(* IEC 61131-3 sources: deprecated-refusr-repo/GP/Main/samples (part 20) *)

(* ---- RND-EXPR_cribs-hyena-lilts.st ---- *)
(*
This code implements a randomly grown symbolic expression:

IN28 & IN39

*)

FUNCTION_BLOCK F_CollectInput
  VAR_IN_OUT
      Data : ARRAY[1..50] OF BOOL;
  END_VAR
  VAR_INPUT
      TICK  : BOOL := 0;
      IN1   : BOOL := 0;
      IN2   : BOOL := 0;
      IN3   : BOOL := 0;
      IN4   : BOOL := 0;
      IN5   : BOOL := 0;
      RESET : BOOL := FALSE;
  END_VAR
  VAR_OUTPUT
      Finished : BOOL;
  END_VAR
  VAR
      j    : USINT := 1;
      tock : BOOL  := 0;
  END_VAR
  IF NOT RESET AND tock = NOT TICK THEN
      Data[j]   := IN1;
      Data[j+1] := IN2;
      Data[j+2] := IN3;
      Data[j+3] := IN4;
      Data[j+4] := IN5;
      j := j + 5;
      tock := TICK;
  ELSE
      j := 1;
      tock := 0;
  END_IF;
  Finished := (j > 50);
END_FUNCTION_BLOCK

PROGRAM Boiler
  VAR
    Data  : ARRAY[1..50] OF BOOL;
    Ready : BOOL;
    CollectInput : F_CollectInput;
  END_VAR
  VAR
    TICK     AT %IX1.0 : BOOL;
    IN1      AT %IX0.3 : BOOL;
    IN2      AT %IX0.4 : BOOL;
    IN3      AT %IX0.5 : BOOL;
    IN4      AT %IX0.6 : BOOL;
    IN5      AT %IX0.7 : BOOL;
    OutReady AT %QX0.0 : BOOL := FALSE;
    FeedNext AT %QX0.1 : BOOL := FALSE;
    Out      AT %QX0.2 : BOOL;
  END_VAR
  CollectInput(TICK:=TICK, IN1:=IN1, IN2:=IN2, IN3:=IN3, IN4:=IN4, IN5:=IN5);
  Ready := CollectInput.Finished;
  FeedNext := 1;
  IF Ready THEN
    Out := (Data[28] AND Data[39]);
    OutReady := 1;
    CollectInput(RESET:=TRUE);
  END_IF;
END_PROGRAM

CONFIGURATION Config0
  RESOURCE Res0 ON PLC
    TASK task0(INTERVAL := T#20ms,PRIORITY := 0);
    PROGRAM instance0 WITH task0 : Boiler;
  END_RESOURCE
END_CONFIGURATION

(* ---- RND-EXPR_culls-boxes-teats.st ---- *)
(*
This code implements a randomly grown symbolic expression:

xor(xor(xor(xor(!((IN48 | (xor(xor(!(!(IN48)), !(!(xor(xor(IN15 & IN37, IN27 & IN43), xor(xor(IN10, IN50), IN49))))), !((IN7 & (xor(xor(IN34, IN29), IN41))) | ((IN34 & IN45) | (!(IN2))))))) & IN16), IN31), IN38), (IN16 | IN47) & IN28), (((!(IN20)) | ((xor(xor(xor(xor(((IN39 | IN35) | (IN9 & IN43)) & IN46, !((!(IN46)) | (xor(xor(IN5, IN34), IN46)))), (!(IN19 | IN49)) | (!(!(IN22)))), xor(xor(IN13, IN22), ((!(IN35)) & (xor(xor(IN2, IN40), IN38))) & IN43)), IN29)) | (xor(xor(!(!(xor(xor(IN8 | IN20, IN6 | IN40), xor(xor(IN12, IN18), IN33)))), !(((!(IN34)) & IN30) | ((!(IN31)) & (IN36 & IN6)))), (!(IN35)) & true)))) & ((((IN17 | (!(!(IN26 | IN42)))) | (xor(xor(IN44, ((xor(xor(IN13, IN3), IN47)) | (xor(xor(IN10, IN45), IN26))) & (xor(xor(!(IN3), IN34 | true), !(IN45)))), !(IN7 | IN35)))) & ((!(!(xor(xor(IN41 & IN25, xor(xor(IN10, IN9), IN48)), IN39)))) | (xor(xor(((xor(xor(IN22, IN35), IN30)) | (IN30 & IN45)) & ((IN24 | IN15) | IN48), !((xor(xor(IN16, IN5), IN23)) | (!(IN4)))), !((xor(xor(IN38, IN16), IN14)) | IN41))))) | ((IN27 & IN46) & ((xor(xor(!(!(xor(xor(IN29, IN24), IN24))), ((IN29 & IN32) & (IN36 | IN47)) | IN15), !(xor(xor(IN45, IN47 | IN29), xor(false, IN9))))) & (xor(xor(xor(xor((xor(xor(IN29, IN4), IN8)) & (!(IN27)), (xor(xor(IN24, IN23), IN10)) | IN19), (IN35 & IN15) | IN20), IN4 & ((!(IN9)) | (xor(xor(IN12, IN15), IN37)))), !(!(IN3)))))))) & (IN27 | IN9))

*)

FUNCTION_BLOCK F_CollectInput
  VAR_IN_OUT
      Data : ARRAY[1..50] OF BOOL;
  END_VAR
  VAR_INPUT
      TICK  : BOOL := 0;
      IN1   : BOOL := 0;
      IN2   : BOOL := 0;
      IN3   : BOOL := 0;
      IN4   : BOOL := 0;
      IN5   : BOOL := 0;
      RESET : BOOL := FALSE;
  END_VAR
  VAR_OUTPUT
      Finished : BOOL;
  END_VAR
  VAR
      j    : USINT := 1;
      tock : BOOL  := 0;
  END_VAR
  IF NOT RESET AND tock = NOT TICK THEN
      Data[j]   := IN1;
      Data[j+1] := IN2;
      Data[j+2] := IN3;
      Data[j+3] := IN4;
      Data[j+4] := IN5;
      j := j + 5;
      tock := TICK;
  ELSE
      j := 1;
      tock := 0;
  END_IF;
  Finished := (j > 50);
END_FUNCTION_BLOCK

PROGRAM Boiler
  VAR
    Data  : ARRAY[1..50] OF BOOL;
    Ready : BOOL;
    CollectInput : F_CollectInput;
  END_VAR
  VAR
    TICK     AT %IX1.0 : BOOL;
    IN1      AT %IX0.3 : BOOL;
    IN2      AT %IX0.4 : BOOL;
    IN3      AT %IX0.5 : BOOL;
    IN4      AT %IX0.6 : BOOL;
    IN5      AT %IX0.7 : BOOL;
    OutReady AT %QX0.0 : BOOL := FALSE;
    FeedNext AT %QX0.1 : BOOL := FALSE;
    Out      AT %QX0.2 : BOOL;
  END_VAR
  CollectInput(TICK:=TICK, IN1:=IN1, IN2:=IN2, IN3:=IN3, IN4:=IN4, IN5:=IN5);
  Ready := CollectInput.Finished;
  FeedNext := 1;
  IF Ready THEN
    Out := (((((NOT ((Data[48] OR (((NOT (NOT Data[48])) XOR (NOT (NOT (((Data[15] AND Data[37]) XOR (Data[27] AND Data[43])) XOR ((Data[10] XOR Data[50]) XOR Data[49]))))) XOR (NOT ((Data[7] AND ((Data[34] XOR Data[29]) XOR Data[41])) OR ((Data[34] AND Data[45]) OR (NOT Data[2])))))) AND Data[16])) XOR Data[31]) XOR Data[38]) XOR ((Data[16] OR Data[47]) AND Data[28])) XOR ((((NOT Data[20]) OR ((((((((Data[39] OR Data[35]) OR (Data[9] AND Data[43])) AND Data[46]) XOR (NOT ((NOT Data[46]) OR ((Data[5] XOR Data[34]) XOR Data[46])))) XOR ((NOT (Data[19] OR Data[49])) OR (NOT (NOT Data[22])))) XOR ((Data[13] XOR Data[22]) XOR (((NOT Data[35]) AND ((Data[2] XOR Data[40]) XOR Data[38])) AND Data[43]))) XOR Data[29]) OR (((NOT (NOT (((Data[8] OR Data[20]) XOR (Data[6] OR Data[40])) XOR ((Data[12] XOR Data[18]) XOR Data[33])))) XOR (NOT (((NOT Data[34]) AND Data[30]) OR ((NOT Data[31]) AND (Data[36] AND Data[6]))))) XOR ((NOT Data[35]) AND TRUE)))) AND ((((Data[17] OR (NOT (NOT (Data[26] OR Data[42])))) OR ((Data[44] XOR ((((Data[13] XOR Data[3]) XOR Data[47]) OR ((Data[10] XOR Data[45]) XOR Data[26])) AND (((NOT Data[3]) XOR (Data[34] OR TRUE)) XOR (NOT Data[45])))) XOR (NOT (Data[7] OR Data[35])))) AND ((NOT (NOT (((Data[41] AND Data[25]) XOR ((Data[10] XOR Data[9]) XOR Data[48])) XOR Data[39]))) OR ((((((Data[22] XOR Data[35]) XOR Data[30]) OR (Data[30] AND Data[45])) AND ((Data[24] OR Data[15]) OR Data[48])) XOR (NOT (((Data[16] XOR Data[5]) XOR Data[23]) OR (NOT Data[4])))) XOR (NOT (((Data[38] XOR Data[16]) XOR Data[14]) OR Data[41]))))) OR ((Data[27] AND Data[46]) AND ((((NOT (NOT ((Data[29] XOR Data[24]) XOR Data[24]))) XOR (((Data[29] AND Data[32]) AND (Data[36] OR Data[47])) OR Data[15])) XOR (NOT ((Data[45] XOR (Data[47] OR Data[29])) XOR (FALSE XOR Data[9])))) AND (((((((Data[29] XOR Data[4]) XOR Data[8]) AND (NOT Data[27])) XOR (((Data[24] XOR Data[23]) XOR Data[10]) OR Data[19])) XOR ((Data[35] AND Data[15]) OR Data[20])) XOR (Data[4] AND ((NOT Data[9]) OR ((Data[12] XOR Data[15]) XOR Data[37])))) XOR (NOT (NOT Data[3]))))))) AND (Data[27] OR Data[9])));
    OutReady := 1;
    CollectInput(RESET:=TRUE);
  END_IF;
END_PROGRAM

CONFIGURATION Config0
  RESOURCE Res0 ON PLC
    TASK task0(INTERVAL := T#20ms,PRIORITY := 0);
    PROGRAM instance0 WITH task0 : Boiler;
  END_RESOURCE
END_CONFIGURATION

(* ---- RND-EXPR_datum-botch-beams.st ---- *)
(*
This code implements a randomly grown symbolic expression:

(((xor(xor((xor(xor(xor(xor(IN19, (!(IN48 | IN21)) & (!(xor(xor(IN30, IN18), IN5)))), IN21), ((xor(xor(IN23 | IN7, IN44 | IN43), IN28 & IN45)) & ((!(IN4)) | (IN37 | IN4))) | (xor(xor((IN10 | IN19) | (IN27 & IN18), IN45), !(IN41)))), IN21)) & ((((IN36 | false) | ((!(IN22)) | (xor(xor(IN17, IN20), IN45)))) | (((xor(xor(IN40, IN49), IN35)) & (!(IN19))) & (xor(xor(xor(xor(IN32, IN22), IN46), !(IN2)), xor(xor(IN46, IN23), IN28))))) | ((((IN7 & IN47) & (IN5 & IN32)) & ((IN29 | IN13) | (true & IN42))) & ((true & (IN8 & IN29)) & (xor(xor(!(IN46), !(IN24)), xor(xor(IN6, IN16), IN4)))))), (((!(!(IN20 | IN46))) | (!(xor(xor(!(IN16), xor(xor(IN12, IN9), IN4)), IN31 | IN40)))) & IN49) & (xor(xor(IN41, (xor(xor((xor(xor(true, IN18), false)) & (xor(xor(IN10, IN15), IN4)), (!(IN14)) & IN12), (IN43 | IN32) & IN32)) & (IN31 | ((xor(xor(IN22, true), IN17)) | (xor(xor(IN49, IN20), false))))), xor(xor(!(IN45), IN46), IN2 | (xor(xor(IN11, IN2 & IN18), IN43 | IN11)))))), IN11)) | IN13) | (xor(xor(xor(xor((!((!((IN29 | IN7) & (IN48 | IN42))) | IN20)) | (!(IN21)), (xor(xor(xor(xor(xor(xor((xor(xor(IN1, IN10), IN29)) | (IN2 & IN25), xor(xor(xor(xor(IN34, IN6), IN25), IN41 & IN10), IN36 & IN25)), (IN6 & IN20) | (IN47 | IN26)), IN7), !((IN43 & IN25) | (xor(xor(IN44, IN44), IN30)))), IN15 | (IN8 & (xor(xor(xor(xor(IN3, IN16), IN33), IN3 & IN40), !(IN40))))), IN31 & IN19)) & (IN27 & (!(IN47 & (xor(xor(IN5, IN38 & IN40), IN30)))))), xor(xor(((!(!(IN24))) & (xor(xor(IN30, IN2), xor(xor(xor(xor(IN38, true), IN8), IN33 & IN9), xor(xor(IN49, IN40), IN43))))) & (((true & (xor(xor(IN49, IN36), IN7))) | ((!(IN21)) | (IN4 & IN40))) & IN47), ((((IN13 | IN3) & IN30) & (xor(xor(IN3 & IN14, !(IN41)), !(IN22)))) & ((!(IN33 | IN21)) | (!(IN18 & IN42)))) | (xor(xor((xor(xor(!(IN37), IN49 | IN14), IN42)) & (!(IN1 & IN30)), ((!(IN18)) & (xor(xor(IN28, IN28), IN42))) & (IN40 | IN32)), !(IN34 & (xor(xor(IN45, IN21), IN18)))))), xor(xor(!(!(xor(xor(IN48 | IN1, !(IN12)), !(IN27)))), ((xor(xor(IN43 | IN15, IN9 | IN20), xor(xor(IN4, IN4), IN11))) & IN35) & (IN21 | (!(IN13 & IN21)))), ((xor(xor(xor(xor(IN29, IN17), IN6), IN23 | IN2), IN46 | IN28)) & (!(IN42))) | IN9))), xor(xor(IN21, !(!(!(!((xor(xor(IN47, IN29), IN31)) & (IN3 & IN43)))))), (!((xor(xor(!(IN27 | IN39), xor(xor(xor(xor(IN1, IN14), IN16), false | IN8), IN47 | IN1)), xor(xor(IN36 & IN31, !(IN39)), IN44 | IN33))) & ((IN8 | (IN5 | IN34)) & (!(xor(xor(IN12, IN31), IN12)))))) | ((((!(xor(xor(IN45, IN8), IN46))) & IN45) & IN8) | (!(!((IN28 & IN42) & (IN50 | IN35))))))), xor(xor(IN29, !((IN34 | (IN1 | (IN12 & (IN6 | IN15)))) & ((!(!(IN32 & IN18))) & (!(!(IN6 & IN28)))))), ((!(!(IN25))) | (xor(xor(xor(xor(!(IN3 & IN34), xor(xor(IN16 & IN26, !(IN26)), IN17)), (IN33 & IN37) & (!(IN32))), ((IN38 | IN8) & (!(IN19))) | (xor(xor(!(IN29), IN4 | IN21), IN39 & IN36))), (xor(xor(IN41 | IN43, xor(xor(IN32, IN10), IN28)), IN18 & IN1)) | (IN25 & IN34)))) & IN8)))) | IN13

*)

FUNCTION_BLOCK F_CollectInput
  VAR_IN_OUT
      Data : ARRAY[1..50] OF BOOL;
  END_VAR
  VAR_INPUT
      TICK  : BOOL := 0;
      IN1   : BOOL := 0;
      IN2   : BOOL := 0;
      IN3   : BOOL := 0;
      IN4   : BOOL := 0;
      IN5   : BOOL := 0;
      RESET : BOOL := FALSE;
  END_VAR
  VAR_OUTPUT
      Finished : BOOL;
  END_VAR
  VAR
      j    : USINT := 1;
      tock : BOOL  := 0;
  END_VAR
  IF NOT RESET AND tock = NOT TICK THEN
      Data[j]   := IN1;
      Data[j+1] := IN2;
      Data[j+2] := IN3;
      Data[j+3] := IN4;
      Data[j+4] := IN5;
      j := j + 5;
      tock := TICK;
  ELSE
      j := 1;
      tock := 0;
  END_IF;
  Finished := (j > 50);
END_FUNCTION_BLOCK

PROGRAM Boiler
  VAR
    Data  : ARRAY[1..50] OF BOOL;
    Ready : BOOL;
    CollectInput : F_CollectInput;
  END_VAR
  VAR
    TICK     AT %IX1.0 : BOOL;
    IN1      AT %IX0.3 : BOOL;
    IN2      AT %IX0.4 : BOOL;
    IN3      AT %IX0.5 : BOOL;
    IN4      AT %IX0.6 : BOOL;
    IN5      AT %IX0.7 : BOOL;
    OutReady AT %QX0.0 : BOOL := FALSE;
    FeedNext AT %QX0.1 : BOOL := FALSE;
    Out      AT %QX0.2 : BOOL;
  END_VAR
  CollectInput(TICK:=TICK, IN1:=IN1, IN2:=IN2, IN3:=IN3, IN4:=IN4, IN5:=IN5);
  Ready := CollectInput.Finished;
  FeedNext := 1;
  IF Ready THEN
    Out := ((((((((((Data[19] XOR ((NOT (Data[48] OR Data[21])) AND (NOT ((Data[30] XOR Data[18]) XOR Data[5])))) XOR Data[21]) XOR (((((Data[23] OR Data[7]) XOR (Data[44] OR Data[43])) XOR (Data[28] AND Data[45])) AND ((NOT Data[4]) OR (Data[37] OR Data[4]))) OR ((((Data[10] OR Data[19]) OR (Data[27] AND Data[18])) XOR Data[45]) XOR (NOT Data[41])))) XOR Data[21]) AND ((((Data[36] OR FALSE) OR ((NOT Data[22]) OR ((Data[17] XOR Data[20]) XOR Data[45]))) OR ((((Data[40] XOR Data[49]) XOR Data[35]) AND (NOT Data[19])) AND ((((Data[32] XOR Data[22]) XOR Data[46]) XOR (NOT Data[2])) XOR ((Data[46] XOR Data[23]) XOR Data[28])))) OR ((((Data[7] AND Data[47]) AND (Data[5] AND Data[32])) AND ((Data[29] OR Data[13]) OR (TRUE AND Data[42]))) AND ((TRUE AND (Data[8] AND Data[29])) AND (((NOT Data[46]) XOR (NOT Data[24])) XOR ((Data[6] XOR Data[16]) XOR Data[4])))))) XOR ((((NOT (NOT (Data[20] OR Data[46]))) OR (NOT (((NOT Data[16]) XOR ((Data[12] XOR Data[9]) XOR Data[4])) XOR (Data[31] OR Data[40])))) AND Data[49]) AND ((Data[41] XOR ((((((TRUE XOR Data[18]) XOR FALSE) AND ((Data[10] XOR Data[15]) XOR Data[4])) XOR ((NOT Data[14]) AND Data[12])) XOR ((Data[43] OR Data[32]) AND Data[32])) AND (Data[31] OR (((Data[22] XOR TRUE) XOR Data[17]) OR ((Data[49] XOR Data[20]) XOR FALSE))))) XOR (((NOT Data[45]) XOR Data[46]) XOR (Data[2] OR ((Data[11] XOR (Data[2] AND Data[18])) XOR (Data[43] OR Data[11]))))))) XOR Data[11]) OR Data[13]) OR ((((((NOT ((NOT ((Data[29] OR Data[7]) AND (Data[48] OR Data[42]))) OR Data[20])) OR (NOT Data[21])) XOR ((((((((((Data[1] XOR Data[10]) XOR Data[29]) OR (Data[2] AND Data[25])) XOR ((((Data[34] XOR Data[6]) XOR Data[25]) XOR (Data[41] AND Data[10])) XOR (Data[36] AND Data[25]))) XOR ((Data[6] AND Data[20]) OR (Data[47] OR Data[26]))) XOR Data[7]) XOR (NOT ((Data[43] AND Data[25]) OR ((Data[44] XOR Data[44]) XOR Data[30])))) XOR (Data[15] OR (Data[8] AND ((((Data[3] XOR Data[16]) XOR Data[33]) XOR (Data[3] AND Data[40])) XOR (NOT Data[40]))))) XOR (Data[31] AND Data[19])) AND (Data[27] AND (NOT (Data[47] AND ((Data[5] XOR (Data[38] AND Data[40])) XOR Data[30])))))) XOR (((((NOT (NOT Data[24])) AND ((Data[30] XOR Data[2]) XOR ((((Data[38] XOR TRUE) XOR Data[8]) XOR (Data[33] AND Data[9])) XOR ((Data[49] XOR Data[40]) XOR Data[43])))) AND (((TRUE AND ((Data[49] XOR Data[36]) XOR Data[7])) OR ((NOT Data[21]) OR (Data[4] AND Data[40]))) AND Data[47])) XOR (((((Data[13] OR Data[3]) AND Data[30]) AND (((Data[3] AND Data[14]) XOR (NOT Data[41])) XOR (NOT Data[22]))) AND ((NOT (Data[33] OR Data[21])) OR (NOT (Data[18] AND Data[42])))) OR ((((((NOT Data[37]) XOR (Data[49] OR Data[14])) XOR Data[42]) AND (NOT (Data[1] AND Data[30]))) XOR (((NOT Data[18]) AND ((Data[28] XOR Data[28]) XOR Data[42])) AND (Data[40] OR Data[32]))) XOR (NOT (Data[34] AND ((Data[45] XOR Data[21]) XOR Data[18])))))) XOR (((NOT (NOT (((Data[48] OR Data[1]) XOR (NOT Data[12])) XOR (NOT Data[27])))) XOR (((((Data[43] OR Data[15]) XOR (Data[9] OR Data[20])) XOR ((Data[4] XOR Data[4]) XOR Data[11])) AND Data[35]) AND (Data[21] OR (NOT (Data[13] AND Data[21]))))) XOR ((((((Data[29] XOR Data[17]) XOR Data[6]) XOR (Data[23] OR Data[2])) XOR (Data[46] OR Data[28])) AND (NOT Data[42])) OR Data[9])))) XOR ((Data[21] XOR (NOT (NOT (NOT (NOT (((Data[47] XOR Data[29]) XOR Data[31]) AND (Data[3] AND Data[43]))))))) XOR ((NOT ((((NOT (Data[27] OR Data[39])) XOR ((((Data[1] XOR Data[14]) XOR Data[16]) XOR (FALSE OR Data[8])) XOR (Data[47] OR Data[1]))) XOR (((Data[36] AND Data[31]) XOR (NOT Data[39])) XOR (Data[44] OR Data[33]))) AND ((Data[8] OR (Data[5] OR Data[34])) AND (NOT ((Data[12] XOR Data[31]) XOR Data[12]))))) OR ((((NOT ((Data[45] XOR Data[8]) XOR Data[46])) AND Data[45]) AND Data[8]) OR (NOT (NOT ((Data[28] AND Data[42]) AND (Data[50] OR Data[35])))))))) XOR ((Data[29] XOR (NOT ((Data[34] OR (Data[1] OR (Data[12] AND (Data[6] OR Data[15])))) AND ((NOT (NOT (Data[32] AND Data[18]))) AND (NOT (NOT (Data[6] AND Data[28]))))))) XOR (((NOT (NOT Data[25])) OR (((((NOT (Data[3] AND Data[34])) XOR (((Data[16] AND Data[26]) XOR (NOT Data[26])) XOR Data[17])) XOR ((Data[33] AND Data[37]) AND (NOT Data[32]))) XOR (((Data[38] OR Data[8]) AND (NOT Data[19])) OR (((NOT Data[29]) XOR (Data[4] OR Data[21])) XOR (Data[39] AND Data[36])))) XOR ((((Data[41] OR Data[43]) XOR ((Data[32] XOR Data[10]) XOR Data[28])) XOR (Data[18] AND Data[1])) OR (Data[25] AND Data[34])))) AND Data[8])))) OR Data[13]);
    OutReady := 1;
    CollectInput(RESET:=TRUE);
  END_IF;
END_PROGRAM

CONFIGURATION Config0
  RESOURCE Res0 ON PLC
    TASK task0(INTERVAL := T#20ms,PRIORITY := 0);
    PROGRAM instance0 WITH task0 : Boiler;
  END_RESOURCE
END_CONFIGURATION

(* ---- RND-EXPR_didot-crows-snoot.st ---- *)
(*
This code implements a randomly grown symbolic expression:

((((xor(xor(IN5, xor(xor(xor(xor(((IN48 & IN29) | (IN9 | IN16)) & ((!(IN32)) & (xor(xor(IN31, IN7), IN31))), IN21 & (!(!(IN38)))), IN40 & ((IN8 & IN7) & (!(IN26)))), !(xor(xor(!(!(IN18)), xor(xor(IN2 & IN4, xor(xor(IN20, IN39), IN3)), IN20)), !(xor(xor(IN38, IN20), IN30))))), xor(xor(!(IN10), xor(xor(IN9, (!(IN6)) & (true & IN13)), xor(xor(xor(xor(IN27, IN43), false), xor(xor(IN49, IN1), IN26)), !(IN6)))), (!(!(IN27))) | (IN47 & (IN34 & IN35))))), (xor(xor(IN44, (!(!(IN15))) & (xor(xor(IN27 & IN46, IN40 & IN32), !(IN14)))), xor(xor(!(IN46 & IN21), !(!(IN46))), (xor(xor(IN25, IN12), IN13)) | (!(IN50))))) | (IN20 | ((!(xor(xor(IN22, IN46), IN28))) | (!(IN24)))))) & (((((IN24 & (!(IN48))) & (!(IN22))) | (!(!(!(IN24))))) | ((xor(xor((!(IN2)) | (!(IN5)), IN46), xor(xor(IN45 & IN25, IN43), IN43))) & (xor(xor(xor(xor(IN7, !(IN33)), xor(xor(IN3, IN5), IN17)), xor(xor(IN39 & IN18, !(IN8)), IN15 & IN24)), (!(IN38)) | (IN9 | IN17))))) & (xor(xor(IN20 & (xor(xor((IN35 | IN47) & (xor(xor(IN46, IN9), IN16)), IN17), xor(xor(!(IN14), IN31), !(IN44)))), xor(xor((xor(xor(xor(xor(IN38, IN15), IN25), IN36 & IN30), IN7 & IN34)) | (!(xor(xor(IN31, IN21), IN10))), !(xor(xor(xor(xor(IN47, IN11), IN2), IN25 | IN46), IN10))), IN21)), IN45)))) | (xor(xor(IN46 & (IN16 | (!((IN31 & (!(IN12))) & (!(IN31 & IN34))))), IN43 | ((!((!(IN7 | IN36)) | IN29)) & (!((xor(xor(!(IN39), IN7), xor(xor(IN2, IN38), IN16))) | (xor(xor(IN21 & IN38, IN39 | IN14), IN28 & IN3)))))), !(!(!(IN5 | (!(IN5 & IN46)))))))) & IN50) & IN18

*)

FUNCTION_BLOCK F_CollectInput
  VAR_IN_OUT
      Data : ARRAY[1..50] OF BOOL;
  END_VAR
  VAR_INPUT
      TICK  : BOOL := 0;
      IN1   : BOOL := 0;
      IN2   : BOOL := 0;
      IN3   : BOOL := 0;
      IN4   : BOOL := 0;
      IN5   : BOOL := 0;
      RESET : BOOL := FALSE;
  END_VAR
  VAR_OUTPUT
      Finished : BOOL;
  END_VAR
  VAR
      j    : USINT := 1;
      tock : BOOL  := 0;
  END_VAR
  IF NOT RESET AND tock = NOT TICK THEN
      Data[j]   := IN1;
      Data[j+1] := IN2;
      Data[j+2] := IN3;
      Data[j+3] := IN4;
      Data[j+4] := IN5;
      j := j + 5;
      tock := TICK;
  ELSE
      j := 1;
      tock := 0;
  END_IF;
  Finished := (j > 50);
END_FUNCTION_BLOCK

PROGRAM Boiler
  VAR
    Data  : ARRAY[1..50] OF BOOL;
    Ready : BOOL;
    CollectInput : F_CollectInput;
  END_VAR
  VAR
    TICK     AT %IX1.0 : BOOL;
    IN1      AT %IX0.3 : BOOL;
    IN2      AT %IX0.4 : BOOL;
    IN3      AT %IX0.5 : BOOL;
    IN4      AT %IX0.6 : BOOL;
    IN5      AT %IX0.7 : BOOL;
    OutReady AT %QX0.0 : BOOL := FALSE;
    FeedNext AT %QX0.1 : BOOL := FALSE;
    Out      AT %QX0.2 : BOOL;
  END_VAR
  CollectInput(TICK:=TICK, IN1:=IN1, IN2:=IN2, IN3:=IN3, IN4:=IN4, IN5:=IN5);
  Ready := CollectInput.Finished;
  FeedNext := 1;
  IF Ready THEN
    Out := ((((((Data[5] XOR (((((((Data[48] AND Data[29]) OR (Data[9] OR Data[16])) AND ((NOT Data[32]) AND ((Data[31] XOR Data[7]) XOR Data[31]))) XOR (Data[21] AND (NOT (NOT Data[38])))) XOR (Data[40] AND ((Data[8] AND Data[7]) AND (NOT Data[26])))) XOR (NOT (((NOT (NOT Data[18])) XOR (((Data[2] AND Data[4]) XOR ((Data[20] XOR Data[39]) XOR Data[3])) XOR Data[20])) XOR (NOT ((Data[38] XOR Data[20]) XOR Data[30]))))) XOR (((NOT Data[10]) XOR ((Data[9] XOR ((NOT Data[6]) AND (TRUE AND Data[13]))) XOR ((((Data[27] XOR Data[43]) XOR FALSE) XOR ((Data[49] XOR Data[1]) XOR Data[26])) XOR (NOT Data[6])))) XOR ((NOT (NOT Data[27])) OR (Data[47] AND (Data[34] AND Data[35])))))) XOR (((Data[44] XOR ((NOT (NOT Data[15])) AND (((Data[27] AND Data[46]) XOR (Data[40] AND Data[32])) XOR (NOT Data[14])))) XOR (((NOT (Data[46] AND Data[21])) XOR (NOT (NOT Data[46]))) XOR (((Data[25] XOR Data[12]) XOR Data[13]) OR (NOT Data[50])))) OR (Data[20] OR ((NOT ((Data[22] XOR Data[46]) XOR Data[28])) OR (NOT Data[24]))))) AND (((((Data[24] AND (NOT Data[48])) AND (NOT Data[22])) OR (NOT (NOT (NOT Data[24])))) OR (((((NOT Data[2]) OR (NOT Data[5])) XOR Data[46]) XOR (((Data[45] AND Data[25]) XOR Data[43]) XOR Data[43])) AND ((((Data[7] XOR (NOT Data[33])) XOR ((Data[3] XOR Data[5]) XOR Data[17])) XOR (((Data[39] AND Data[18]) XOR (NOT Data[8])) XOR (Data[15] AND Data[24]))) XOR ((NOT Data[38]) OR (Data[9] OR Data[17]))))) AND (((Data[20] AND ((((Data[35] OR Data[47]) AND ((Data[46] XOR Data[9]) XOR Data[16])) XOR Data[17]) XOR (((NOT Data[14]) XOR Data[31]) XOR (NOT Data[44])))) XOR (((((((Data[38] XOR Data[15]) XOR Data[25]) XOR (Data[36] AND Data[30])) XOR (Data[7] AND Data[34])) OR (NOT ((Data[31] XOR Data[21]) XOR Data[10]))) XOR (NOT ((((Data[47] XOR Data[11]) XOR Data[2]) XOR (Data[25] OR Data[46])) XOR Data[10]))) XOR Data[21])) XOR Data[45]))) OR (((Data[46] AND (Data[16] OR (NOT ((Data[31] AND (NOT Data[12])) AND (NOT (Data[31] AND Data[34])))))) XOR (Data[43] OR ((NOT ((NOT (Data[7] OR Data[36])) OR Data[29])) AND (NOT ((((NOT Data[39]) XOR Data[7]) XOR ((Data[2] XOR Data[38]) XOR Data[16])) OR (((Data[21] AND Data[38]) XOR (Data[39] OR Data[14])) XOR (Data[28] AND Data[3]))))))) XOR (NOT (NOT (NOT (Data[5] OR (NOT (Data[5] AND Data[46])))))))) AND Data[50]) AND Data[18]);
    OutReady := 1;
    CollectInput(RESET:=TRUE);
  END_IF;
END_PROGRAM

CONFIGURATION Config0
  RESOURCE Res0 ON PLC
    TASK task0(INTERVAL := T#20ms,PRIORITY := 0);
    PROGRAM instance0 WITH task0 : Boiler;
  END_RESOURCE
END_CONFIGURATION

(* ---- RND-EXPR_dotty-douse-lurer.st ---- *)
(*
This code implements a randomly grown symbolic expression:

xor(xor(!(xor(xor(((xor(xor(IN28, false), (xor(xor((IN5 | IN20) & IN27, (IN25 & IN12) & (!(IN47))), xor(xor(IN14 | IN16, xor(xor(IN17, IN42), IN9)), IN6 | IN50))) | (!(xor(xor(IN20 & IN18, IN41 & false), !(IN41)))))) & (!(!(xor(xor((IN4 | IN22) | (IN4 & IN4), (!(IN31)) & (!(IN11))), !(!(IN25))))))) | (IN22 | (!((((IN15 | IN11) & (IN10 | IN33)) | ((xor(xor(IN28, IN28), IN26)) & (IN10 & IN11))) | IN27))), !(!((xor(xor((xor(xor(IN4 & IN11, xor(xor(IN28, IN40), IN2)), IN2 | IN17)) & (!(IN16)), xor(xor(IN21 | (IN43 | IN19), xor(xor(IN42, IN25 | IN18), IN25 & IN49)), xor(xor(true, IN35 | true), !(IN36)))), (!(IN6 & IN31)) | (!(IN42 & IN48)))) & (xor(xor(IN22, (!(IN30)) | (xor(xor(!(IN11), !(IN42)), IN1 | IN27))), IN7 | ((IN2 | IN23) | (IN30 | IN49))))))), !(IN20 | (IN16 & ((!((IN39 & IN22) & (!(IN7)))) | (!(xor(xor(IN8 | IN15, IN21 | IN44), !(IN2))))))))), IN28), !(!(IN41 | (!(xor(xor(!(xor(xor(xor(xor(IN34 | IN30, IN36), xor(xor(IN31, IN38), IN14)), xor(xor(IN7 & IN44, IN11 & IN13), IN5 & IN15)), !(IN11 & IN10))), (IN14 | false) | IN29), (!(IN47)) & (!((xor(xor(IN17, IN6), IN4)) | (IN47 | IN10)))))))))

*)

FUNCTION_BLOCK F_CollectInput
  VAR_IN_OUT
      Data : ARRAY[1..50] OF BOOL;
  END_VAR
  VAR_INPUT
      TICK  : BOOL := 0;
      IN1   : BOOL := 0;
      IN2   : BOOL := 0;
      IN3   : BOOL := 0;
      IN4   : BOOL := 0;
      IN5   : BOOL := 0;
      RESET : BOOL := FALSE;
  END_VAR
  VAR_OUTPUT
      Finished : BOOL;
  END_VAR
  VAR
      j    : USINT := 1;
      tock : BOOL  := 0;
  END_VAR
  IF NOT RESET AND tock = NOT TICK THEN
      Data[j]   := IN1;
      Data[j+1] := IN2;
      Data[j+2] := IN3;
      Data[j+3] := IN4;
      Data[j+4] := IN5;
      j := j + 5;
      tock := TICK;
  ELSE
      j := 1;
      tock := 0;
  END_IF;
  Finished := (j > 50);
END_FUNCTION_BLOCK

PROGRAM Boiler
  VAR
    Data  : ARRAY[1..50] OF BOOL;
    Ready : BOOL;
    CollectInput : F_CollectInput;
  END_VAR
  VAR
    TICK     AT %IX1.0 : BOOL;
    IN1      AT %IX0.3 : BOOL;
    IN2      AT %IX0.4 : BOOL;
    IN3      AT %IX0.5 : BOOL;
    IN4      AT %IX0.6 : BOOL;
    IN5      AT %IX0.7 : BOOL;
    OutReady AT %QX0.0 : BOOL := FALSE;
    FeedNext AT %QX0.1 : BOOL := FALSE;
    Out      AT %QX0.2 : BOOL;
  END_VAR
  CollectInput(TICK:=TICK, IN1:=IN1, IN2:=IN2, IN3:=IN3, IN4:=IN4, IN5:=IN5);
  Ready := CollectInput.Finished;
  FeedNext := 1;
  IF Ready THEN
    Out := (((NOT ((((((Data[28] XOR FALSE) XOR (((((Data[5] OR Data[20]) AND Data[27]) XOR ((Data[25] AND Data[12]) AND (NOT Data[47]))) XOR (((Data[14] OR Data[16]) XOR ((Data[17] XOR Data[42]) XOR Data[9])) XOR (Data[6] OR Data[50]))) OR (NOT (((Data[20] AND Data[18]) XOR (Data[41] AND FALSE)) XOR (NOT Data[41]))))) AND (NOT (NOT ((((Data[4] OR Data[22]) OR (Data[4] AND Data[4])) XOR ((NOT Data[31]) AND (NOT Data[11]))) XOR (NOT (NOT Data[25])))))) OR (Data[22] OR (NOT ((((Data[15] OR Data[11]) AND (Data[10] OR Data[33])) OR (((Data[28] XOR Data[28]) XOR Data[26]) AND (Data[10] AND Data[11]))) OR Data[27])))) XOR (NOT (NOT (((((((Data[4] AND Data[11]) XOR ((Data[28] XOR Data[40]) XOR Data[2])) XOR (Data[2] OR Data[17])) AND (NOT Data[16])) XOR (((Data[21] OR (Data[43] OR Data[19])) XOR ((Data[42] XOR (Data[25] OR Data[18])) XOR (Data[25] AND Data[49]))) XOR ((TRUE XOR (Data[35] OR TRUE)) XOR (NOT Data[36])))) XOR ((NOT (Data[6] AND Data[31])) OR (NOT (Data[42] AND Data[48])))) AND ((Data[22] XOR ((NOT Data[30]) OR (((NOT Data[11]) XOR (NOT Data[42])) XOR (Data[1] OR Data[27])))) XOR (Data[7] OR ((Data[2] OR Data[23]) OR (Data[30] OR Data[49])))))))) XOR (NOT (Data[20] OR (Data[16] AND ((NOT ((Data[39] AND Data[22]) AND (NOT Data[7]))) OR (NOT (((Data[8] OR Data[15]) XOR (Data[21] OR Data[44])) XOR (NOT Data[2]))))))))) XOR Data[28]) XOR (NOT (NOT (Data[41] OR (NOT (((NOT (((((Data[34] OR Data[30]) XOR Data[36]) XOR ((Data[31] XOR Data[38]) XOR Data[14])) XOR (((Data[7] AND Data[44]) XOR (Data[11] AND Data[13])) XOR (Data[5] AND Data[15]))) XOR (NOT (Data[11] AND Data[10])))) XOR ((Data[14] OR FALSE) OR Data[29])) XOR ((NOT Data[47]) AND (NOT (((Data[17] XOR Data[6]) XOR Data[4]) OR (Data[47] OR Data[10]))))))))));
    OutReady := 1;
    CollectInput(RESET:=TRUE);
  END_IF;
END_PROGRAM

CONFIGURATION Config0
  RESOURCE Res0 ON PLC
    TASK task0(INTERVAL := T#20ms,PRIORITY := 0);
    PROGRAM instance0 WITH task0 : Boiler;
  END_RESOURCE
END_CONFIGURATION

(* ---- RND-EXPR_doxie-capos-donna.st ---- *)
(*
This code implements a randomly grown symbolic expression:

!(!(xor(xor(IN7 | ((((!(xor(xor(IN46, IN6 & IN48), IN36 | IN35))) | (!((xor(xor(IN26, IN22), IN45)) | (IN5 | true)))) | (!(((IN23 & IN25) & IN7) | (xor(xor(xor(xor(IN6, IN4), true), xor(xor(IN2, IN20), IN9)), xor(xor(IN4, IN11), IN36)))))) & (!(IN23))), IN8), ((!((((IN36 & IN24) | (IN45 | IN45)) | ((!(IN8)) | (!(IN23)))) & ((xor(xor(xor(xor(IN41, IN42), IN5), xor(xor(IN5, IN3), IN41)), xor(xor(IN20, IN39), true))) & (xor(xor(!(IN12), IN47 & false), IN14 & IN23))))) | (xor(xor((!(IN3)) & (((xor(xor(IN24, IN43), IN28)) | (!(IN10))) & (!(IN22 | IN28))), IN16), (xor(xor(IN1, IN1), (IN16 & true) | (IN40 | IN50))) & (!(IN39 & (IN8 & IN8)))))) | IN3)))

*)

FUNCTION_BLOCK F_CollectInput
  VAR_IN_OUT
      Data : ARRAY[1..50] OF BOOL;
  END_VAR
  VAR_INPUT
      TICK  : BOOL := 0;
      IN1   : BOOL := 0;
      IN2   : BOOL := 0;
      IN3   : BOOL := 0;
      IN4   : BOOL := 0;
      IN5   : BOOL := 0;
      RESET : BOOL := FALSE;
  END_VAR
  VAR_OUTPUT
      Finished : BOOL;
  END_VAR
  VAR
      j    : USINT := 1;
      tock : BOOL  := 0;
  END_VAR
  IF NOT RESET AND tock = NOT TICK THEN
      Data[j]   := IN1;
      Data[j+1] := IN2;
      Data[j+2] := IN3;
      Data[j+3] := IN4;
      Data[j+4] := IN5;
      j := j + 5;
      tock := TICK;
  ELSE
      j := 1;
      tock := 0;
  END_IF;
  Finished := (j > 50);
END_FUNCTION_BLOCK

PROGRAM Boiler
  VAR
    Data  : ARRAY[1..50] OF BOOL;
    Ready : BOOL;
    CollectInput : F_CollectInput;
  END_VAR
  VAR
    TICK     AT %IX1.0 : BOOL;
    IN1      AT %IX0.3 : BOOL;
    IN2      AT %IX0.4 : BOOL;
    IN3      AT %IX0.5 : BOOL;
    IN4      AT %IX0.6 : BOOL;
    IN5      AT %IX0.7 : BOOL;
    OutReady AT %QX0.0 : BOOL := FALSE;
    FeedNext AT %QX0.1 : BOOL := FALSE;
    Out      AT %QX0.2 : BOOL;
  END_VAR
  CollectInput(TICK:=TICK, IN1:=IN1, IN2:=IN2, IN3:=IN3, IN4:=IN4, IN5:=IN5);
  Ready := CollectInput.Finished;
  FeedNext := 1;
  IF Ready THEN
    Out := (NOT (NOT (((Data[7] OR ((((NOT ((Data[46] XOR (Data[6] AND Data[48])) XOR (Data[36] OR Data[35]))) OR (NOT (((Data[26] XOR Data[22]) XOR Data[45]) OR (Data[5] OR TRUE)))) OR (NOT (((Data[23] AND Data[25]) AND Data[7]) OR ((((Data[6] XOR Data[4]) XOR TRUE) XOR ((Data[2] XOR Data[20]) XOR Data[9])) XOR ((Data[4] XOR Data[11]) XOR Data[36]))))) AND (NOT Data[23]))) XOR Data[8]) XOR (((NOT ((((Data[36] AND Data[24]) OR (Data[45] OR Data[45])) OR ((NOT Data[8]) OR (NOT Data[23]))) AND (((((Data[41] XOR Data[42]) XOR Data[5]) XOR ((Data[5] XOR Data[3]) XOR Data[41])) XOR ((Data[20] XOR Data[39]) XOR TRUE)) AND (((NOT Data[12]) XOR (Data[47] AND FALSE)) XOR (Data[14] AND Data[23]))))) OR ((((NOT Data[3]) AND ((((Data[24] XOR Data[43]) XOR Data[28]) OR (NOT Data[10])) AND (NOT (Data[22] OR Data[28])))) XOR Data[16]) XOR (((Data[1] XOR Data[1]) XOR ((Data[16] AND TRUE) OR (Data[40] OR Data[50]))) AND (NOT (Data[39] AND (Data[8] AND Data[8])))))) OR Data[3]))));
    OutReady := 1;
    CollectInput(RESET:=TRUE);
  END_IF;
END_PROGRAM

CONFIGURATION Config0
  RESOURCE Res0 ON PLC
    TASK task0(INTERVAL := T#20ms,PRIORITY := 0);
    PROGRAM instance0 WITH task0 : Boiler;
  END_RESOURCE
END_CONFIGURATION

(* ---- RND-EXPR_dungs-zesty-molar.st ---- *)
(*
This code implements a randomly grown symbolic expression:

!(((xor(xor(IN8, IN20), IN48)) & ((xor(xor(IN35, (xor(xor(IN29, IN4), xor(xor(xor(xor(IN24, IN13 & IN7), IN43 & IN37), xor(xor(IN22 | IN45, !(IN45)), IN29)), (IN25 | IN31) & (!(IN35))))) & ((!(IN17)) | (!(!(!(IN20)))))), (xor(xor(xor(xor((!(IN19)) & (xor(xor(IN33, IN6), true)), (IN15 | IN42) | (!(IN44))), (xor(xor(IN21, IN29), IN28)) | (xor(xor(IN7, IN40), IN24))), IN25), xor(xor(!(xor(xor(IN31, IN7), IN47)), (IN19 & IN22) & (xor(xor(IN43, IN25), IN31))), !(xor(xor(IN50, IN27), IN7))))) | IN38)) | (((!(!((IN47 & false) & (IN22 | IN14)))) & (xor(xor((IN36 & (xor(xor(IN24, IN34), IN34))) | ((IN28 & IN4) | (xor(xor(IN18, IN20), IN30))), (xor(xor(xor(xor(IN31, IN19), IN48), IN44 & IN44), IN23 | IN36)) & ((!(IN27)) & IN36)), !(xor(xor(xor(xor(IN25, IN47), IN30), IN48 & IN3), IN37))))) & IN1))) | (IN9 | IN17))

*)

FUNCTION_BLOCK F_CollectInput
  VAR_IN_OUT
      Data : ARRAY[1..50] OF BOOL;
  END_VAR
  VAR_INPUT
      TICK  : BOOL := 0;
      IN1   : BOOL := 0;
      IN2   : BOOL := 0;
      IN3   : BOOL := 0;
      IN4   : BOOL := 0;
      IN5   : BOOL := 0;
      RESET : BOOL := FALSE;
  END_VAR
  VAR_OUTPUT
      Finished : BOOL;
  END_VAR
  VAR
      j    : USINT := 1;
      tock : BOOL  := 0;
  END_VAR
  IF NOT RESET AND tock = NOT TICK THEN
      Data[j]   := IN1;
      Data[j+1] := IN2;
      Data[j+2] := IN3;
      Data[j+3] := IN4;
      Data[j+4] := IN5;
      j := j + 5;
      tock := TICK;
  ELSE
      j := 1;
      tock := 0;
  END_IF;
  Finished := (j > 50);
END_FUNCTION_BLOCK

PROGRAM Boiler
  VAR
    Data  : ARRAY[1..50] OF BOOL;
    Ready : BOOL;
    CollectInput : F_CollectInput;
  END_VAR
  VAR
    TICK     AT %IX1.0 : BOOL;
    IN1      AT %IX0.3 : BOOL;
    IN2      AT %IX0.4 : BOOL;
    IN3      AT %IX0.5 : BOOL;
    IN4      AT %IX0.6 : BOOL;
    IN5      AT %IX0.7 : BOOL;
    OutReady AT %QX0.0 : BOOL := FALSE;
    FeedNext AT %QX0.1 : BOOL := FALSE;
    Out      AT %QX0.2 : BOOL;
  END_VAR
  CollectInput(TICK:=TICK, IN1:=IN1, IN2:=IN2, IN3:=IN3, IN4:=IN4, IN5:=IN5);
  Ready := CollectInput.Finished;
  FeedNext := 1;
  IF Ready THEN
    Out := (NOT ((((Data[8] XOR Data[20]) XOR Data[48]) AND (((Data[35] XOR (((Data[29] XOR Data[4]) XOR ((((Data[24] XOR (Data[13] AND Data[7])) XOR (Data[43] AND Data[37])) XOR (((Data[22] OR Data[45]) XOR (NOT Data[45])) XOR Data[29])) XOR ((Data[25] OR Data[31]) AND (NOT Data[35])))) AND ((NOT Data[17]) OR (NOT (NOT (NOT Data[20])))))) XOR (((((((NOT Data[19]) AND ((Data[33] XOR Data[6]) XOR TRUE)) XOR ((Data[15] OR Data[42]) OR (NOT Data[44]))) XOR (((Data[21] XOR Data[29]) XOR Data[28]) OR ((Data[7] XOR Data[40]) XOR Data[24]))) XOR Data[25]) XOR (((NOT ((Data[31] XOR Data[7]) XOR Data[47])) XOR ((Data[19] AND Data[22]) AND ((Data[43] XOR Data[25]) XOR Data[31]))) XOR (NOT ((Data[50] XOR Data[27]) XOR Data[7])))) OR Data[38])) OR (((NOT (NOT ((Data[47] AND FALSE) AND (Data[22] OR Data[14])))) AND ((((Data[36] AND ((Data[24] XOR Data[34]) XOR Data[34])) OR ((Data[28] AND Data[4]) OR ((Data[18] XOR Data[20]) XOR Data[30]))) XOR (((((Data[31] XOR Data[19]) XOR Data[48]) XOR (Data[44] AND Data[44])) XOR (Data[23] OR Data[36])) AND ((NOT Data[27]) AND Data[36]))) XOR (NOT ((((Data[25] XOR Data[47]) XOR Data[30]) XOR (Data[48] AND Data[3])) XOR Data[37])))) AND Data[1]))) OR (Data[9] OR Data[17])));
    OutReady := 1;
    CollectInput(RESET:=TRUE);
  END_IF;
END_PROGRAM

CONFIGURATION Config0
  RESOURCE Res0 ON PLC
    TASK task0(INTERVAL := T#20ms,PRIORITY := 0);
    PROGRAM instance0 WITH task0 : Boiler;
  END_RESOURCE
END_CONFIGURATION

(* ---- RND-EXPR_eagle-ingot-brawn.st ---- *)
(*
This code implements a randomly grown symbolic expression:

(IN32 & (xor(xor((!(IN11 | ((xor(xor(IN13, !(IN3 | IN42)), !(IN34))) & IN11))) | ((!((((IN19 | IN12) & (xor(xor(IN42, IN27), IN13))) & ((!(IN24)) | (!(IN42)))) & (!(IN16)))) & IN2), ((xor(xor((xor(xor((IN17 & IN7) & (xor(xor(IN27, IN22), true)), (xor(xor(true, IN43), IN46)) | IN50), IN7)) & ((xor(xor(IN42, xor(xor(IN25, IN34), IN24)), !(IN12))) & ((IN7 | IN34) & (!(IN30)))), (xor(xor(IN14, !(IN8 | IN22)), (!(IN18)) & IN38)) & (((!(IN1)) | (!(IN7))) & ((IN10 & IN17) | false))), xor(xor(!(IN46), xor(xor((IN29 & IN48) & IN38, (xor(xor(IN11, IN9), IN22)) | (xor(xor(IN45, IN16), IN44))), (!(IN25)) | IN37)), !(xor(xor(!(IN18), xor(xor(IN29, IN45), IN27)), IN36 | IN6))))) & ((!(xor(xor(xor(xor(!(IN42), !(IN45)), xor(xor(IN2, IN30), IN11)), xor(xor(IN13 & false, IN1 & IN37), IN38 | IN33)), xor(xor(xor(xor(IN49, IN40), IN47), IN36), true)))) & ((xor(xor(xor(xor(IN35, !(IN29)), IN30), IN3), IN47 & (xor(xor(IN32, IN25), IN23)))) & (xor(xor((IN20 | IN24) & (!(IN4)), !(IN4)), (IN24 | IN5) & (IN50 | IN29)))))) | IN32), !(IN27)))) | (((!(IN34)) | ((xor(xor(((((xor(xor(IN43, IN35), IN19)) & IN1) | ((IN26 | IN10) | (IN1 & IN49))) & ((IN33 | (IN43 | IN37)) & IN42)) & ((!((IN13 | IN6) & (xor(xor(IN22, IN43), IN26)))) & (((xor(xor(IN48, IN4), IN6)) & IN39) & (!(IN17 & false)))), xor(xor(((!(!(IN12))) | IN38) & (xor(xor((IN42 & IN23) & (IN5 | IN11), xor(xor(IN28 & true, IN15), !(IN24))), (xor(xor(IN14, IN19), IN43)) | (!(IN18)))), (!(xor(xor(IN48, IN46 | IN20), !(IN37)))) | (xor(xor(IN7 | (IN16 & IN40), (xor(xor(IN30, IN26), IN26)) | (false & IN24)), (!(IN29)) & IN23))), IN12 & (!(IN37)))), ((xor(xor(xor(xor(IN5 & IN19, IN23), !(IN27)), IN23), (IN9 | IN49) | (!(IN44)))) & (!(xor(xor(!(IN34), IN4), xor(xor(false, IN6), IN47))))) | (xor(xor(xor(xor(IN10 | (!(IN13)), IN14), !(IN48 & IN32)), xor(xor(IN29, xor(xor(IN46 | IN14, IN18), IN49 & IN49)), false)), IN23 | IN23)))) & (xor(xor((xor(xor(!(xor(xor(xor(xor(IN33, IN36), IN5), IN13 & true), IN35 | IN17)), !((!(IN16)) | (xor(xor(IN3, IN11), true)))), (xor(xor(xor(xor(IN47, IN50), false), IN9 & IN29), xor(xor(IN17, IN40), IN9))) & (xor(xor(xor(xor(IN48, IN21), IN13), IN47 | IN38), IN5 | IN26)))) & IN19, IN40), !(((!(IN22 | IN28)) & ((xor(xor(IN46, IN22), IN38)) & IN20)) & (!((!(IN48)) & (IN46 & IN40)))))))) | ((!(!(IN27))) & (((!(xor(xor(IN11, xor(xor(xor(xor(xor(xor(IN22, IN25), IN30), xor(xor(IN6, IN26), IN21)), !(IN45)), xor(xor(xor(xor(IN38, IN43), IN33), IN38 & IN39), IN26 | IN30)), (IN31 | IN47) & (IN30 & IN35))), ((!(IN9)) | IN41) | ((IN19 | IN40) & (!(IN37)))))) & IN38) | IN19)))

*)

FUNCTION_BLOCK F_CollectInput
  VAR_IN_OUT
      Data : ARRAY[1..50] OF BOOL;
  END_VAR
  VAR_INPUT
      TICK  : BOOL := 0;
      IN1   : BOOL := 0;
      IN2   : BOOL := 0;
      IN3   : BOOL := 0;
      IN4   : BOOL := 0;
      IN5   : BOOL := 0;
      RESET : BOOL := FALSE;
  END_VAR
  VAR_OUTPUT
      Finished : BOOL;
  END_VAR
  VAR
      j    : USINT := 1;
      tock : BOOL  := 0;
  END_VAR
  IF NOT RESET AND tock = NOT TICK THEN
      Data[j]   := IN1;
      Data[j+1] := IN2;
      Data[j+2] := IN3;
      Data[j+3] := IN4;
      Data[j+4] := IN5;
      j := j + 5;
      tock := TICK;
  ELSE
      j := 1;
      tock := 0;
  END_IF;
  Finished := (j > 50);
END_FUNCTION_BLOCK

PROGRAM Boiler
  VAR
    Data  : ARRAY[1..50] OF BOOL;
    Ready : BOOL;
    CollectInput : F_CollectInput;
  END_VAR
  VAR
    TICK     AT %IX1.0 : BOOL;
    IN1      AT %IX0.3 : BOOL;
    IN2      AT %IX0.4 : BOOL;
    IN3      AT %IX0.5 : BOOL;
    IN4      AT %IX0.6 : BOOL;
    IN5      AT %IX0.7 : BOOL;
    OutReady AT %QX0.0 : BOOL := FALSE;
    FeedNext AT %QX0.1 : BOOL := FALSE;
    Out      AT %QX0.2 : BOOL;
  END_VAR
  CollectInput(TICK:=TICK, IN1:=IN1, IN2:=IN2, IN3:=IN3, IN4:=IN4, IN5:=IN5);
  Ready := CollectInput.Finished;
  FeedNext := 1;
  IF Ready THEN
    Out := ((Data[32] AND ((((NOT (Data[11] OR (((Data[13] XOR (NOT (Data[3] OR Data[42]))) XOR (NOT Data[34])) AND Data[11]))) OR ((NOT ((((Data[19] OR Data[12]) AND ((Data[42] XOR Data[27]) XOR Data[13])) AND ((NOT Data[24]) OR (NOT Data[42]))) AND (NOT Data[16]))) AND Data[2])) XOR (((((((((Data[17] AND Data[7]) AND ((Data[27] XOR Data[22]) XOR TRUE)) XOR (((TRUE XOR Data[43]) XOR Data[46]) OR Data[50])) XOR Data[7]) AND (((Data[42] XOR ((Data[25] XOR Data[34]) XOR Data[24])) XOR (NOT Data[12])) AND ((Data[7] OR Data[34]) AND (NOT Data[30])))) XOR (((Data[14] XOR (NOT (Data[8] OR Data[22]))) XOR ((NOT Data[18]) AND Data[38])) AND (((NOT Data[1]) OR (NOT Data[7])) AND ((Data[10] AND Data[17]) OR FALSE)))) XOR (((NOT Data[46]) XOR ((((Data[29] AND Data[48]) AND Data[38]) XOR (((Data[11] XOR Data[9]) XOR Data[22]) OR ((Data[45] XOR Data[16]) XOR Data[44]))) XOR ((NOT Data[25]) OR Data[37]))) XOR (NOT (((NOT Data[18]) XOR ((Data[29] XOR Data[45]) XOR Data[27])) XOR (Data[36] OR Data[6]))))) AND ((NOT (((((NOT Data[42]) XOR (NOT Data[45])) XOR ((Data[2] XOR Data[30]) XOR Data[11])) XOR (((Data[13] AND FALSE) XOR (Data[1] AND Data[37])) XOR (Data[38] OR Data[33]))) XOR ((((Data[49] XOR Data[40]) XOR Data[47]) XOR Data[36]) XOR TRUE))) AND (((((Data[35] XOR (NOT Data[29])) XOR Data[30]) XOR Data[3]) XOR (Data[47] AND ((Data[32] XOR Data[25]) XOR Data[23]))) AND ((((Data[20] OR Data[24]) AND (NOT Data[4])) XOR (NOT Data[4])) XOR ((Data[24] OR Data[5]) AND (Data[50] OR Data[29])))))) OR Data[32])) XOR (NOT Data[27]))) OR (((NOT Data[34]) OR (((((((((Data[43] XOR Data[35]) XOR Data[19]) AND Data[1]) OR ((Data[26] OR Data[10]) OR (Data[1] AND Data[49]))) AND ((Data[33] OR (Data[43] OR Data[37])) AND Data[42])) AND ((NOT ((Data[13] OR Data[6]) AND ((Data[22] XOR Data[43]) XOR Data[26]))) AND ((((Data[48] XOR Data[4]) XOR Data[6]) AND Data[39]) AND (NOT (Data[17] AND FALSE))))) XOR (((((NOT (NOT Data[12])) OR Data[38]) AND ((((Data[42] AND Data[23]) AND (Data[5] OR Data[11])) XOR (((Data[28] AND TRUE) XOR Data[15]) XOR (NOT Data[24]))) XOR (((Data[14] XOR Data[19]) XOR Data[43]) OR (NOT Data[18])))) XOR ((NOT ((Data[48] XOR (Data[46] OR Data[20])) XOR (NOT Data[37]))) OR (((Data[7] OR (Data[16] AND Data[40])) XOR (((Data[30] XOR Data[26]) XOR Data[26]) OR (FALSE AND Data[24]))) XOR ((NOT Data[29]) AND Data[23])))) XOR (Data[12] AND (NOT Data[37])))) XOR (((((((Data[5] AND Data[19]) XOR Data[23]) XOR (NOT Data[27])) XOR Data[23]) XOR ((Data[9] OR Data[49]) OR (NOT Data[44]))) AND (NOT (((NOT Data[34]) XOR Data[4]) XOR ((FALSE XOR Data[6]) XOR Data[47])))) OR (((((Data[10] OR (NOT Data[13])) XOR Data[14]) XOR (NOT (Data[48] AND Data[32]))) XOR ((Data[29] XOR (((Data[46] OR Data[14]) XOR Data[18]) XOR (Data[49] AND Data[49]))) XOR FALSE)) XOR (Data[23] OR Data[23])))) AND ((((((NOT ((((Data[33] XOR Data[36]) XOR Data[5]) XOR (Data[13] AND TRUE)) XOR (Data[35] OR Data[17]))) XOR (NOT ((NOT Data[16]) OR ((Data[3] XOR Data[11]) XOR TRUE)))) XOR (((((Data[47] XOR Data[50]) XOR FALSE) XOR (Data[9] AND Data[29])) XOR ((Data[17] XOR Data[40]) XOR Data[9])) AND ((((Data[48] XOR Data[21]) XOR Data[13]) XOR (Data[47] OR Data[38])) XOR (Data[5] OR Data[26])))) AND Data[19]) XOR Data[40]) XOR (NOT (((NOT (Data[22] OR Data[28])) AND (((Data[46] XOR Data[22]) XOR Data[38]) AND Data[20])) AND (NOT ((NOT Data[48]) AND (Data[46] AND Data[40])))))))) OR ((NOT (NOT Data[27])) AND (((NOT ((Data[11] XOR ((((((Data[22] XOR Data[25]) XOR Data[30]) XOR ((Data[6] XOR Data[26]) XOR Data[21])) XOR (NOT Data[45])) XOR ((((Data[38] XOR Data[43]) XOR Data[33]) XOR (Data[38] AND Data[39])) XOR (Data[26] OR Data[30]))) XOR ((Data[31] OR Data[47]) AND (Data[30] AND Data[35])))) XOR (((NOT Data[9]) OR Data[41]) OR ((Data[19] OR Data[40]) AND (NOT Data[37]))))) AND Data[38]) OR Data[19]))));
    OutReady := 1;
    CollectInput(RESET:=TRUE);
  END_IF;
END_PROGRAM

CONFIGURATION Config0
  RESOURCE Res0 ON PLC
    TASK task0(INTERVAL := T#20ms,PRIORITY := 0);
    PROGRAM instance0 WITH task0 : Boiler;
  END_RESOURCE
END_CONFIGURATION

(* ---- RND-EXPR_emote-trout-maybe.st ---- *)
(*
This code implements a randomly grown symbolic expression:

!(!(((xor(xor(xor(xor((((xor(xor(IN1, IN36), IN46)) & IN23) | IN28) | (((!(IN17)) & (xor(xor(IN44, IN26), IN12))) | (!(IN13 & IN19))), IN10), !(IN20)), !(!(!(xor(xor(IN46, IN23 & IN30), IN17 & IN43))))), IN6 | IN14)) | ((!(IN14)) | (!(xor(xor(xor(xor(!(!(IN5)), IN33 & (!(IN16))), (xor(xor(IN28, IN38), IN24)) | (!(IN44))), ((xor(xor(IN27, IN29), IN10)) | (IN42 & IN46)) | (!(IN20 | IN29))), !(!(xor(xor(IN43, IN36), IN42)))))))) & IN24))

*)

FUNCTION_BLOCK F_CollectInput
  VAR_IN_OUT
      Data : ARRAY[1..50] OF BOOL;
  END_VAR
  VAR_INPUT
      TICK  : BOOL := 0;
      IN1   : BOOL := 0;
      IN2   : BOOL := 0;
      IN3   : BOOL := 0;
      IN4   : BOOL := 0;
      IN5   : BOOL := 0;
      RESET : BOOL := FALSE;
  END_VAR
  VAR_OUTPUT
      Finished : BOOL;
  END_VAR
  VAR
      j    : USINT := 1;
      tock : BOOL  := 0;
  END_VAR
  IF NOT RESET AND tock = NOT TICK THEN
      Data[j]   := IN1;
      Data[j+1] := IN2;
      Data[j+2] := IN3;
      Data[j+3] := IN4;
      Data[j+4] := IN5;
      j := j + 5;
      tock := TICK;
  ELSE
      j := 1;
      tock := 0;
  END_IF;
  Finished := (j > 50);
END_FUNCTION_BLOCK

PROGRAM Boiler
  VAR
    Data  : ARRAY[1..50] OF BOOL;
    Ready : BOOL;
    CollectInput : F_CollectInput;
  END_VAR
  VAR
    TICK     AT %IX1.0 : BOOL;
    IN1      AT %IX0.3 : BOOL;
    IN2      AT %IX0.4 : BOOL;
    IN3      AT %IX0.5 : BOOL;
    IN4      AT %IX0.6 : BOOL;
    IN5      AT %IX0.7 : BOOL;
    OutReady AT %QX0.0 : BOOL := FALSE;
    FeedNext AT %QX0.1 : BOOL := FALSE;
    Out      AT %QX0.2 : BOOL;
  END_VAR
  CollectInput(TICK:=TICK, IN1:=IN1, IN2:=IN2, IN3:=IN3, IN4:=IN4, IN5:=IN5);
  Ready := CollectInput.Finished;
  FeedNext := 1;
  IF Ready THEN
    Out := (NOT (NOT (((((((((((Data[1] XOR Data[36]) XOR Data[46]) AND Data[23]) OR Data[28]) OR (((NOT Data[17]) AND ((Data[44] XOR Data[26]) XOR Data[12])) OR (NOT (Data[13] AND Data[19])))) XOR Data[10]) XOR (NOT Data[20])) XOR (NOT (NOT (NOT ((Data[46] XOR (Data[23] AND Data[30])) XOR (Data[17] AND Data[43])))))) XOR (Data[6] OR Data[14])) OR ((NOT Data[14]) OR (NOT (((((NOT (NOT Data[5])) XOR (Data[33] AND (NOT Data[16]))) XOR (((Data[28] XOR Data[38]) XOR Data[24]) OR (NOT Data[44]))) XOR ((((Data[27] XOR Data[29]) XOR Data[10]) OR (Data[42] AND Data[46])) OR (NOT (Data[20] OR Data[29])))) XOR (NOT (NOT ((Data[43] XOR Data[36]) XOR Data[42]))))))) AND Data[24])));
    OutReady := 1;
    CollectInput(RESET:=TRUE);
  END_IF;
END_PROGRAM

CONFIGURATION Config0
  RESOURCE Res0 ON PLC
    TASK task0(INTERVAL := T#20ms,PRIORITY := 0);
    PROGRAM instance0 WITH task0 : Boiler;
  END_RESOURCE
END_CONFIGURATION

(* ---- RND-EXPR_eruct-dorks-laird.st ---- *)
(*
This code implements a randomly grown symbolic expression:

(IN21 & (xor(xor(((IN15 | (xor(xor(((xor(xor(IN46, IN46), IN48)) & (IN48 & IN37)) | (xor(xor(IN13 & IN17, IN18 | IN36), IN43)), (!(IN20 & IN16)) & (true & IN10)), xor(xor((IN8 & IN24) & (IN6 | IN40), (IN20 | IN43) & (!(IN22))), IN27 & (IN16 & IN29))))) | (IN7 & IN37)) | ((xor(xor(IN49, IN22), ((!(!(IN10))) & IN12) & (((IN2 | IN15) | (IN30 | IN34)) | (!(IN42 & IN45))))) & ((!(xor(xor(IN33 & IN39, (IN12 & IN13) & (IN8 | IN38)), (!(IN4)) | (!(IN49))))) | (!(!((IN44 | IN30) & IN11))))), xor(xor(((!(xor(xor(IN49 | (IN16 | IN40), (IN21 | IN13) & IN42), !(IN49 & IN21)))) | IN48) | (xor(xor(IN9, (((IN32 | IN17) & (!(IN31))) & ((!(IN28)) & (IN43 | IN29))) & (true & ((xor(xor(false, IN29), IN12)) & (IN14 & IN39)))), !(!(xor(xor(IN17, !(IN48)), IN15 & IN25))))), IN29), (((xor(xor(xor(xor(IN40, IN33 & IN22), IN31 | IN14), IN27), (!(IN9)) & (xor(xor(IN25, IN49), IN10)))) | ((xor(xor(!(IN2), IN1), IN6 & IN12)) | IN35)) | ((xor(xor(IN27, !(!(IN28))), IN33)) & (!((!(IN11)) | (!(IN46)))))) | (xor(xor(IN28, IN39), !(xor(xor(!(IN49), xor(xor(xor(xor(IN46, IN9), IN37), IN36), IN35 | IN27)), xor(xor(IN8 | IN24, IN20 & IN28), IN20))))))), IN25))) & IN46

*)

FUNCTION_BLOCK F_CollectInput
  VAR_IN_OUT
      Data : ARRAY[1..50] OF BOOL;
  END_VAR
  VAR_INPUT
      TICK  : BOOL := 0;
      IN1   : BOOL := 0;
      IN2   : BOOL := 0;
      IN3   : BOOL := 0;
      IN4   : BOOL := 0;
      IN5   : BOOL := 0;
      RESET : BOOL := FALSE;
  END_VAR
  VAR_OUTPUT
      Finished : BOOL;
  END_VAR
  VAR
      j    : USINT := 1;
      tock : BOOL  := 0;
  END_VAR
  IF NOT RESET AND tock = NOT TICK THEN
      Data[j]   := IN1;
      Data[j+1] := IN2;
      Data[j+2] := IN3;
      Data[j+3] := IN4;
      Data[j+4] := IN5;
      j := j + 5;
      tock := TICK;
  ELSE
      j := 1;
      tock := 0;
  END_IF;
  Finished := (j > 50);
END_FUNCTION_BLOCK

PROGRAM Boiler
  VAR
    Data  : ARRAY[1..50] OF BOOL;
    Ready : BOOL;
    CollectInput : F_CollectInput;
  END_VAR
  VAR
    TICK     AT %IX1.0 : BOOL;
    IN1      AT %IX0.3 : BOOL;
    IN2      AT %IX0.4 : BOOL;
    IN3      AT %IX0.5 : BOOL;
    IN4      AT %IX0.6 : BOOL;
    IN5      AT %IX0.7 : BOOL;
    OutReady AT %QX0.0 : BOOL := FALSE;
    FeedNext AT %QX0.1 : BOOL := FALSE;
    Out      AT %QX0.2 : BOOL;
  END_VAR
  CollectInput(TICK:=TICK, IN1:=IN1, IN2:=IN2, IN3:=IN3, IN4:=IN4, IN5:=IN5);
  Ready := CollectInput.Finished;
  FeedNext := 1;
  IF Ready THEN
    Out := ((Data[21] AND (((((Data[15] OR ((((((Data[46] XOR Data[46]) XOR Data[48]) AND (Data[48] AND Data[37])) OR (((Data[13] AND Data[17]) XOR (Data[18] OR Data[36])) XOR Data[43])) XOR ((NOT (Data[20] AND Data[16])) AND (TRUE AND Data[10]))) XOR ((((Data[8] AND Data[24]) AND (Data[6] OR Data[40])) XOR ((Data[20] OR Data[43]) AND (NOT Data[22]))) XOR (Data[27] AND (Data[16] AND Data[29]))))) OR (Data[7] AND Data[37])) OR (((Data[49] XOR Data[22]) XOR (((NOT (NOT Data[10])) AND Data[12]) AND (((Data[2] OR Data[15]) OR (Data[30] OR Data[34])) OR (NOT (Data[42] AND Data[45]))))) AND ((NOT (((Data[33] AND Data[39]) XOR ((Data[12] AND Data[13]) AND (Data[8] OR Data[38]))) XOR ((NOT Data[4]) OR (NOT Data[49])))) OR (NOT (NOT ((Data[44] OR Data[30]) AND Data[11])))))) XOR (((((NOT (((Data[49] OR (Data[16] OR Data[40])) XOR ((Data[21] OR Data[13]) AND Data[42])) XOR (NOT (Data[49] AND Data[21])))) OR Data[48]) OR ((Data[9] XOR ((((Data[32] OR Data[17]) AND (NOT Data[31])) AND ((NOT Data[28]) AND (Data[43] OR Data[29]))) AND (TRUE AND (((FALSE XOR Data[29]) XOR Data[12]) AND (Data[14] AND Data[39]))))) XOR (NOT (NOT ((Data[17] XOR (NOT Data[48])) XOR (Data[15] AND Data[25])))))) XOR Data[29]) XOR (((((((Data[40] XOR (Data[33] AND Data[22])) XOR (Data[31] OR Data[14])) XOR Data[27]) XOR ((NOT Data[9]) AND ((Data[25] XOR Data[49]) XOR Data[10]))) OR ((((NOT Data[2]) XOR Data[1]) XOR (Data[6] AND Data[12])) OR Data[35])) OR (((Data[27] XOR (NOT (NOT Data[28]))) XOR Data[33]) AND (NOT ((NOT Data[11]) OR (NOT Data[46]))))) OR ((Data[28] XOR Data[39]) XOR (NOT (((NOT Data[49]) XOR ((((Data[46] XOR Data[9]) XOR Data[37]) XOR Data[36]) XOR (Data[35] OR Data[27]))) XOR (((Data[8] OR Data[24]) XOR (Data[20] AND Data[28])) XOR Data[20]))))))) XOR Data[25])) AND Data[46]);
    OutReady := 1;
    CollectInput(RESET:=TRUE);
  END_IF;
END_PROGRAM

CONFIGURATION Config0
  RESOURCE Res0 ON PLC
    TASK task0(INTERVAL := T#20ms,PRIORITY := 0);
    PROGRAM instance0 WITH task0 : Boiler;
  END_RESOURCE
END_CONFIGURATION

(* ---- RND-EXPR_fleas-nooky-enema.st ---- *)
(*
This code implements a randomly grown symbolic expression:

!((!(IN47 & (!(IN17 | ((((!(IN4)) & (IN14 | IN5)) | (IN32 & (xor(xor(IN6, IN2), IN30)))) | (((xor(xor(IN35, IN6), IN22)) & (IN2 & IN10)) & ((xor(xor(IN5, IN30), IN41)) | (xor(xor(IN25, IN3), IN21))))))))) | (((xor(xor(IN27 & (!(!(IN12 | IN44))), IN27), !(xor(xor(IN48 | (!(false & IN37)), xor(xor((xor(xor(IN27, IN45), IN24)) | (IN16 & IN23), !(IN15)), IN13)), IN9 | (!(!(IN47))))))) & (xor(xor((!(xor(xor(!(IN21), !(IN16)), IN31))) & ((!((!(IN8)) | (IN35 & IN25))) | ((xor(xor(xor(xor(IN48, IN19), IN9), IN8 & IN35), IN45 | IN30)) & ((IN36 | IN34) | (IN29 & IN1)))), !((!((IN24 | IN8) | (xor(xor(IN14, IN34), IN43)))) | ((!(IN24)) & ((IN15 & IN6) | (!(IN20)))))), IN27))) | (xor(xor(IN5, ((((!(xor(xor(IN39, IN37), IN36))) | (xor(xor(xor(xor(IN47, IN13), IN15), IN32 & IN23), !(IN14)))) | (((!(IN26)) | (!(IN36))) | ((IN6 | IN24) & (!(IN33))))) & ((!(xor(xor(IN20 & IN40, xor(xor(IN40, IN32), IN35)), IN5))) | IN22)) & IN40), !(xor(xor(IN49, IN31 & (xor(xor(IN23, xor(xor(xor(xor(IN12, IN22), IN32), IN48), false & IN1)), (IN11 | IN17) | (IN43 | IN11)))), ((xor(xor(xor(xor(IN17, IN20), IN17), IN10 | IN2), IN32 | IN34)) & (!(!(IN34)))) & (((!(IN34)) | (true & IN39)) & ((IN5 | IN6) | (IN44 | IN35)))))))))

*)

FUNCTION_BLOCK F_CollectInput
  VAR_IN_OUT
      Data : ARRAY[1..50] OF BOOL;
  END_VAR
  VAR_INPUT
      TICK  : BOOL := 0;
      IN1   : BOOL := 0;
      IN2   : BOOL := 0;
      IN3   : BOOL := 0;
      IN4   : BOOL := 0;
      IN5   : BOOL := 0;
      RESET : BOOL := FALSE;
  END_VAR
  VAR_OUTPUT
      Finished : BOOL;
  END_VAR
  VAR
      j    : USINT := 1;
      tock : BOOL  := 0;
  END_VAR
  IF NOT RESET AND tock = NOT TICK THEN
      Data[j]   := IN1;
      Data[j+1] := IN2;
      Data[j+2] := IN3;
      Data[j+3] := IN4;
      Data[j+4] := IN5;
      j := j + 5;
      tock := TICK;
  ELSE
      j := 1;
      tock := 0;
  END_IF;
  Finished := (j > 50);
END_FUNCTION_BLOCK

PROGRAM Boiler
  VAR
    Data  : ARRAY[1..50] OF BOOL;
    Ready : BOOL;
    CollectInput : F_CollectInput;
  END_VAR
  VAR
    TICK     AT %IX1.0 : BOOL;
    IN1      AT %IX0.3 : BOOL;
    IN2      AT %IX0.4 : BOOL;
    IN3      AT %IX0.5 : BOOL;
    IN4      AT %IX0.6 : BOOL;
    IN5      AT %IX0.7 : BOOL;
    OutReady AT %QX0.0 : BOOL := FALSE;
    FeedNext AT %QX0.1 : BOOL := FALSE;
    Out      AT %QX0.2 : BOOL;
  END_VAR
  CollectInput(TICK:=TICK, IN1:=IN1, IN2:=IN2, IN3:=IN3, IN4:=IN4, IN5:=IN5);
  Ready := CollectInput.Finished;
  FeedNext := 1;
  IF Ready THEN
    Out := (NOT ((NOT (Data[47] AND (NOT (Data[17] OR ((((NOT Data[4]) AND (Data[14] OR Data[5])) OR (Data[32] AND ((Data[6] XOR Data[2]) XOR Data[30]))) OR ((((Data[35] XOR Data[6]) XOR Data[22]) AND (Data[2] AND Data[10])) AND (((Data[5] XOR Data[30]) XOR Data[41]) OR ((Data[25] XOR Data[3]) XOR Data[21])))))))) OR (((((Data[27] AND (NOT (NOT (Data[12] OR Data[44])))) XOR Data[27]) XOR (NOT (((Data[48] OR (NOT (FALSE AND Data[37]))) XOR (((((Data[27] XOR Data[45]) XOR Data[24]) OR (Data[16] AND Data[23])) XOR (NOT Data[15])) XOR Data[13])) XOR (Data[9] OR (NOT (NOT Data[47])))))) AND ((((NOT (((NOT Data[21]) XOR (NOT Data[16])) XOR Data[31])) AND ((NOT ((NOT Data[8]) OR (Data[35] AND Data[25]))) OR (((((Data[48] XOR Data[19]) XOR Data[9]) XOR (Data[8] AND Data[35])) XOR (Data[45] OR Data[30])) AND ((Data[36] OR Data[34]) OR (Data[29] AND Data[1]))))) XOR (NOT ((NOT ((Data[24] OR Data[8]) OR ((Data[14] XOR Data[34]) XOR Data[43]))) OR ((NOT Data[24]) AND ((Data[15] AND Data[6]) OR (NOT Data[20])))))) XOR Data[27])) OR ((Data[5] XOR (((((NOT ((Data[39] XOR Data[37]) XOR Data[36])) OR ((((Data[47] XOR Data[13]) XOR Data[15]) XOR (Data[32] AND Data[23])) XOR (NOT Data[14]))) OR (((NOT Data[26]) OR (NOT Data[36])) OR ((Data[6] OR Data[24]) AND (NOT Data[33])))) AND ((NOT (((Data[20] AND Data[40]) XOR ((Data[40] XOR Data[32]) XOR Data[35])) XOR Data[5])) OR Data[22])) AND Data[40])) XOR (NOT ((Data[49] XOR (Data[31] AND ((Data[23] XOR ((((Data[12] XOR Data[22]) XOR Data[32]) XOR Data[48]) XOR (FALSE AND Data[1]))) XOR ((Data[11] OR Data[17]) OR (Data[43] OR Data[11]))))) XOR ((((((Data[17] XOR Data[20]) XOR Data[17]) XOR (Data[10] OR Data[2])) XOR (Data[32] OR Data[34])) AND (NOT (NOT Data[34]))) AND (((NOT Data[34]) OR (TRUE AND Data[39])) AND ((Data[5] OR Data[6]) OR (Data[44] OR Data[35]))))))))));
    OutReady := 1;
    CollectInput(RESET:=TRUE);
  END_IF;
END_PROGRAM

CONFIGURATION Config0
  RESOURCE Res0 ON PLC
    TASK task0(INTERVAL := T#20ms,PRIORITY := 0);
    PROGRAM instance0 WITH task0 : Boiler;
  END_RESOURCE
END_CONFIGURATION

(* ---- RND-EXPR_freer-nadir-vague.st ---- *)
(*
This code implements a randomly grown symbolic expression:

(!(((!(((xor(xor(xor(xor(xor(xor(IN30, IN19), IN50), xor(xor(IN35, IN19), IN44)), IN29), !(IN28 & IN18)), xor(xor(IN26 | IN48, !(IN15)), xor(xor(IN24, IN37), IN46)))) & (!((IN8 & IN3) | (!(IN18))))) | ((((IN9 & IN43) & (IN49 | IN43)) | ((!(IN42)) | (IN47 | false))) | IN2))) | (xor(xor(IN16, IN19 & (xor(xor((IN36 & true) | (!(IN22)), xor(xor((!(IN39)) & (!(IN8)), (IN10 | IN24) | (IN5 | IN4)), (!(IN28)) & (IN24 & false))), ((xor(xor(IN6, IN1), IN15)) & (!(IN20))) | ((xor(xor(IN28, IN49), IN12)) & (xor(xor(IN2, IN46), IN24)))))), (IN19 | IN26) & (!((IN3 & (IN8 & IN41)) & (IN31 & (xor(xor(IN5, IN21), IN6)))))))) & (xor(xor(IN12, !((!(IN28 & (!(!(IN23))))) & ((xor(xor(!(!(IN33)), (xor(xor(IN50, IN35), IN39)) & (IN42 & IN32)), false)) | IN2))), ((xor(xor(!(!(IN42 & IN19)), IN45), ((IN22 | IN23) | IN36) | (xor(xor(IN13, IN48 | IN7), IN24 | IN8)))) | (!(!(xor(xor(IN19 | IN14, IN2), !(IN48)))))) & (xor(xor(IN44, IN17), xor(xor(!(!(!(IN36))), xor(xor(xor(xor(IN26 & IN14, IN25 | IN18), IN37), xor(xor(!(IN33), IN25 & false), xor(xor(IN1, IN12), IN4))), !(!(IN22)))), IN3))))))) | (((IN47 | (xor(xor(xor(xor(IN7, IN44), !(IN46)), (xor(xor(IN9, IN46 & (IN31 | (!(IN4)))), true | (IN46 & (xor(xor(IN2, true), IN27))))) | ((!(IN1)) & (((!(IN46)) & (IN19 | IN18)) | ((xor(xor(IN4, IN5), IN25)) | (xor(xor(IN50, IN13), IN33)))))), !((xor(xor(xor(xor(!(IN42), xor(xor(IN10, IN36), true)), IN5 & IN27), xor(xor(IN27 | IN46, xor(xor(IN31, IN5), IN11)), !(IN29))), (xor(xor(IN28, IN9), IN31)) | (xor(xor(IN37, IN32), IN4)))) & IN2)))) | ((xor(xor(IN20, !(xor(xor((xor(xor(IN17 & IN10, xor(xor(IN1, IN35), IN47)), IN12 & IN2)) & (xor(xor(xor(xor(IN4, IN42), IN35), IN23 | IN3), IN37)), IN24), !(xor(xor(IN40, IN29), !(IN21)))))), (IN12 & (xor(xor(IN13, !(IN48)), !(xor(xor(IN19, IN8), IN13))))) | (!(xor(xor(!(IN5 | IN11), (IN26 | IN26) | (xor(xor(IN10, IN49), IN32))), !(!(IN3))))))) | IN12)) & IN35)

*)

FUNCTION_BLOCK F_CollectInput
  VAR_IN_OUT
      Data : ARRAY[1..50] OF BOOL;
  END_VAR
  VAR_INPUT
      TICK  : BOOL := 0;
      IN1   : BOOL := 0;
      IN2   : BOOL := 0;
      IN3   : BOOL := 0;
      IN4   : BOOL := 0;
      IN5   : BOOL := 0;
      RESET : BOOL := FALSE;
  END_VAR
  VAR_OUTPUT
      Finished : BOOL;
  END_VAR
  VAR
      j    : USINT := 1;
      tock : BOOL  := 0;
  END_VAR
  IF NOT RESET AND tock = NOT TICK THEN
      Data[j]   := IN1;
      Data[j+1] := IN2;
      Data[j+2] := IN3;
      Data[j+3] := IN4;
      Data[j+4] := IN5;
      j := j + 5;
      tock := TICK;
  ELSE
      j := 1;
      tock := 0;
  END_IF;
  Finished := (j > 50);
END_FUNCTION_BLOCK

PROGRAM Boiler
  VAR
    Data  : ARRAY[1..50] OF BOOL;
    Ready : BOOL;
    CollectInput : F_CollectInput;
  END_VAR
  VAR
    TICK     AT %IX1.0 : BOOL;
    IN1      AT %IX0.3 : BOOL;
    IN2      AT %IX0.4 : BOOL;
    IN3      AT %IX0.5 : BOOL;
    IN4      AT %IX0.6 : BOOL;
    IN5      AT %IX0.7 : BOOL;
    OutReady AT %QX0.0 : BOOL := FALSE;
    FeedNext AT %QX0.1 : BOOL := FALSE;
    Out      AT %QX0.2 : BOOL;
  END_VAR
  CollectInput(TICK:=TICK, IN1:=IN1, IN2:=IN2, IN3:=IN3, IN4:=IN4, IN5:=IN5);
  Ready := CollectInput.Finished;
  FeedNext := 1;
  IF Ready THEN
    Out := ((NOT (((NOT ((((((((Data[30] XOR Data[19]) XOR Data[50]) XOR ((Data[35] XOR Data[19]) XOR Data[44])) XOR Data[29]) XOR (NOT (Data[28] AND Data[18]))) XOR (((Data[26] OR Data[48]) XOR (NOT Data[15])) XOR ((Data[24] XOR Data[37]) XOR Data[46]))) AND (NOT ((Data[8] AND Data[3]) OR (NOT Data[18])))) OR ((((Data[9] AND Data[43]) AND (Data[49] OR Data[43])) OR ((NOT Data[42]) OR (Data[47] OR FALSE))) OR Data[2]))) OR ((Data[16] XOR (Data[19] AND ((((Data[36] AND TRUE) OR (NOT Data[22])) XOR ((((NOT Data[39]) AND (NOT Data[8])) XOR ((Data[10] OR Data[24]) OR (Data[5] OR Data[4]))) XOR ((NOT Data[28]) AND (Data[24] AND FALSE)))) XOR ((((Data[6] XOR Data[1]) XOR Data[15]) AND (NOT Data[20])) OR (((Data[28] XOR Data[49]) XOR Data[12]) AND ((Data[2] XOR Data[46]) XOR Data[24])))))) XOR ((Data[19] OR Data[26]) AND (NOT ((Data[3] AND (Data[8] AND Data[41])) AND (Data[31] AND ((Data[5] XOR Data[21]) XOR Data[6]))))))) AND ((Data[12] XOR (NOT ((NOT (Data[28] AND (NOT (NOT Data[23])))) AND ((((NOT (NOT Data[33])) XOR (((Data[50] XOR Data[35]) XOR Data[39]) AND (Data[42] AND Data[32]))) XOR FALSE) OR Data[2])))) XOR (((((NOT (NOT (Data[42] AND Data[19]))) XOR Data[45]) XOR (((Data[22] OR Data[23]) OR Data[36]) OR ((Data[13] XOR (Data[48] OR Data[7])) XOR (Data[24] OR Data[8])))) OR (NOT (NOT (((Data[19] OR Data[14]) XOR Data[2]) XOR (NOT Data[48]))))) AND ((Data[44] XOR Data[17]) XOR (((NOT (NOT (NOT Data[36]))) XOR (((((Data[26] AND Data[14]) XOR (Data[25] OR Data[18])) XOR Data[37]) XOR (((NOT Data[33]) XOR (Data[25] AND FALSE)) XOR ((Data[1] XOR Data[12]) XOR Data[4]))) XOR (NOT (NOT Data[22])))) XOR Data[3])))))) OR (((Data[47] OR ((((Data[7] XOR Data[44]) XOR (NOT Data[46])) XOR (((Data[9] XOR (Data[46] AND (Data[31] OR (NOT Data[4])))) XOR (TRUE OR (Data[46] AND ((Data[2] XOR TRUE) XOR Data[27])))) OR ((NOT Data[1]) AND (((NOT Data[46]) AND (Data[19] OR Data[18])) OR (((Data[4] XOR Data[5]) XOR Data[25]) OR ((Data[50] XOR Data[13]) XOR Data[33])))))) XOR (NOT ((((((NOT Data[42]) XOR ((Data[10] XOR Data[36]) XOR TRUE)) XOR (Data[5] AND Data[27])) XOR (((Data[27] OR Data[46]) XOR ((Data[31] XOR Data[5]) XOR Data[11])) XOR (NOT Data[29]))) XOR (((Data[28] XOR Data[9]) XOR Data[31]) OR ((Data[37] XOR Data[32]) XOR Data[4]))) AND Data[2])))) OR (((Data[20] XOR (NOT ((((((Data[17] AND Data[10]) XOR ((Data[1] XOR Data[35]) XOR Data[47])) XOR (Data[12] AND Data[2])) AND ((((Data[4] XOR Data[42]) XOR Data[35]) XOR (Data[23] OR Data[3])) XOR Data[37])) XOR Data[24]) XOR (NOT ((Data[40] XOR Data[29]) XOR (NOT Data[21])))))) XOR ((Data[12] AND ((Data[13] XOR (NOT Data[48])) XOR (NOT ((Data[19] XOR Data[8]) XOR Data[13])))) OR (NOT (((NOT (Data[5] OR Data[11])) XOR ((Data[26] OR Data[26]) OR ((Data[10] XOR Data[49]) XOR Data[32]))) XOR (NOT (NOT Data[3])))))) OR Data[12])) AND Data[35]));
    OutReady := 1;
    CollectInput(RESET:=TRUE);
  END_IF;
END_PROGRAM

CONFIGURATION Config0
  RESOURCE Res0 ON PLC
    TASK task0(INTERVAL := T#20ms,PRIORITY := 0);
    PROGRAM instance0 WITH task0 : Boiler;
  END_RESOURCE
END_CONFIGURATION

(* ---- RND-EXPR_grits-papas-auric.st ---- *)
(*
This code implements a randomly grown symbolic expression:

(xor(xor(IN33, (xor(xor(xor(xor(IN4 | (xor(xor(IN46 | IN42, IN14), xor(xor(xor(xor(IN23, xor(xor(true, IN1), IN23)), !(IN34)), xor(xor(IN49 | IN6, IN44), xor(xor(IN24, IN34), IN27))), (IN2 | IN3) | (!(IN43))))), IN40 | IN3), xor(xor(IN10, IN11 & ((false & IN19) & IN47)), (xor(xor((!(IN28)) & (IN22 & IN37), IN2), xor(xor(IN30 & IN18, IN4 | IN45), IN37 | IN8))) | ((!(!(IN6))) | ((!(IN23)) | (IN26 | IN23))))), IN24 & (((xor(xor(xor(xor(IN30, xor(xor(IN46, IN26), IN48)), IN47 & IN29), (IN1 | IN13) & (!(IN48))), !(IN42 & IN3))) & IN27) | ((!(IN40 & IN46)) & (xor(xor(xor(xor(IN32 | IN26, IN42 & IN6), !(IN28)), !(xor(xor(true, IN50), IN22))), IN47 | (!(IN32))))))), (!(((xor(xor(IN46 | IN26, IN10), IN37 & IN14)) & (!(xor(xor(IN31, IN18), IN21)))) & IN28)) & (IN10 & (xor(xor(IN6 | (xor(xor(IN42, xor(xor(IN40, IN44), IN19)), IN48)), xor(xor(xor(xor(!(IN35), xor(xor(IN9, IN11), IN20)), xor(xor(IN50, IN25), IN1)), IN6 | (xor(xor(IN9, IN18), IN18))), xor(xor(IN44 & IN22, !(IN9)), IN25))), IN26 & IN38))))) | (xor(xor(true & ((xor(xor((!(IN23 | IN16)) & (!(xor(xor(IN22, IN50), IN9))), (xor(xor(!(IN42), !(IN14)), xor(xor(IN3, IN34), IN28))) | (!(!(IN24)))), (IN25 & (IN40 & IN13)) & (IN5 | (xor(xor(IN10, IN1), IN31))))) & ((xor(xor(!(IN8 & IN33), (xor(xor(IN17, IN34), IN34)) & IN6), (xor(xor(IN7, IN43), IN13)) & IN11)) | (xor(xor(IN34, !(xor(xor(IN41, true), IN49))), (xor(xor(IN39, IN49), IN43)) & (xor(xor(IN30, IN26), IN36)))))), IN41 & (((((IN18 | false) & (IN50 | IN45)) | (xor(xor(IN9 | IN7, !(IN18)), IN34 | IN21))) & IN6) | (xor(xor(IN40, xor(xor(IN7, false), (IN17 & IN37) & IN24)), (!(IN16)) | (!(IN22 | IN8)))))), IN16))), IN9 | (!(xor(xor(IN8, (!((xor(xor(IN18 | IN28, IN17 & IN6), true | IN4)) | (!(xor(xor(IN26, IN22), IN30))))) | (xor(xor((!(IN4)) & (xor(xor(IN48 | IN34, IN39 | IN15), IN41 & IN46)), !(!(!(IN32)))), xor(xor(!(!(IN13)), IN23), IN8)))), xor(xor(IN9, (IN35 & (IN3 & (IN43 | IN44))) & (IN21 | (IN3 & (xor(xor(IN4, IN50), IN21))))), xor(xor(xor(xor(IN29 & (!(IN40)), xor(xor(IN32 & IN21, IN10 & IN25), xor(xor(false, IN32), IN24))), !(IN18 & IN45)), (IN46 & (IN27 & IN23)) | IN3), xor(xor(!(IN32 | IN3), (IN48 & IN28) | (IN18 & IN4)), xor(xor(IN38 & IN23, !(IN48)), IN1))))))))) | (!((((xor(xor(IN14 | (xor(xor(!(IN18 & IN27), (!(IN46)) | (!(IN22))), (!(IN15)) | (xor(xor(IN27, IN25), IN25)))), xor(xor(xor(xor(xor(xor(xor(xor(IN48, IN20), IN49), !(IN6)), IN21 | IN24), !(xor(xor(IN45, IN13), IN7))), !(IN16)), xor(xor((IN41 | IN27) & (IN19 & IN19), IN46), IN49)), !(IN3))), IN6)) | (IN18 & ((xor(xor((IN35 & IN46) | (IN19 | IN12), !(xor(xor(IN35, IN22), IN28))), (IN36 & IN18) | (!(IN43)))) & ((xor(xor(xor(xor(IN40, IN26), IN18), IN33 & IN31), !(IN43))) & (xor(xor(IN5 | IN20, IN36), xor(xor(IN18, IN49), IN12))))))) | IN26) & IN18))

*)

FUNCTION_BLOCK F_CollectInput
  VAR_IN_OUT
      Data : ARRAY[1..50] OF BOOL;
  END_VAR
  VAR_INPUT
      TICK  : BOOL := 0;
      IN1   : BOOL := 0;
      IN2   : BOOL := 0;
      IN3   : BOOL := 0;
      IN4   : BOOL := 0;
      IN5   : BOOL := 0;
      RESET : BOOL := FALSE;
  END_VAR
  VAR_OUTPUT
      Finished : BOOL;
  END_VAR
  VAR
      j    : USINT := 1;
      tock : BOOL  := 0;
  END_VAR
  IF NOT RESET AND tock = NOT TICK THEN
      Data[j]   := IN1;
      Data[j+1] := IN2;
      Data[j+2] := IN3;
      Data[j+3] := IN4;
      Data[j+4] := IN5;
      j := j + 5;
      tock := TICK;
  ELSE
      j := 1;
      tock := 0;
  END_IF;
  Finished := (j > 50);
END_FUNCTION_BLOCK

PROGRAM Boiler
  VAR
    Data  : ARRAY[1..50] OF BOOL;
    Ready : BOOL;
    CollectInput : F_CollectInput;
  END_VAR
  VAR
    TICK     AT %IX1.0 : BOOL;
    IN1      AT %IX0.3 : BOOL;
    IN2      AT %IX0.4 : BOOL;
    IN3      AT %IX0.5 : BOOL;
    IN4      AT %IX0.6 : BOOL;
    IN5      AT %IX0.7 : BOOL;
    OutReady AT %QX0.0 : BOOL := FALSE;
    FeedNext AT %QX0.1 : BOOL := FALSE;
    Out      AT %QX0.2 : BOOL;
  END_VAR
  CollectInput(TICK:=TICK, IN1:=IN1, IN2:=IN2, IN3:=IN3, IN4:=IN4, IN5:=IN5);
  Ready := CollectInput.Finished;
  FeedNext := 1;
  IF Ready THEN
    Out := (((Data[33] XOR ((((((Data[4] OR (((Data[46] OR Data[42]) XOR Data[14]) XOR ((((Data[23] XOR ((TRUE XOR Data[1]) XOR Data[23])) XOR (NOT Data[34])) XOR (((Data[49] OR Data[6]) XOR Data[44]) XOR ((Data[24] XOR Data[34]) XOR Data[27]))) XOR ((Data[2] OR Data[3]) OR (NOT Data[43]))))) XOR (Data[40] OR Data[3])) XOR ((Data[10] XOR (Data[11] AND ((FALSE AND Data[19]) AND Data[47]))) XOR (((((NOT Data[28]) AND (Data[22] AND Data[37])) XOR Data[2]) XOR (((Data[30] AND Data[18]) XOR (Data[4] OR Data[45])) XOR (Data[37] OR Data[8]))) OR ((NOT (NOT Data[6])) OR ((NOT Data[23]) OR (Data[26] OR Data[23])))))) XOR (Data[24] AND ((((((Data[30] XOR ((Data[46] XOR Data[26]) XOR Data[48])) XOR (Data[47] AND Data[29])) XOR ((Data[1] OR Data[13]) AND (NOT Data[48]))) XOR (NOT (Data[42] AND Data[3]))) AND Data[27]) OR ((NOT (Data[40] AND Data[46])) AND (((((Data[32] OR Data[26]) XOR (Data[42] AND Data[6])) XOR (NOT Data[28])) XOR (NOT ((TRUE XOR Data[50]) XOR Data[22]))) XOR (Data[47] OR (NOT Data[32]))))))) XOR ((NOT (((((Data[46] OR Data[26]) XOR Data[10]) XOR (Data[37] AND Data[14])) AND (NOT ((Data[31] XOR Data[18]) XOR Data[21]))) AND Data[28])) AND (Data[10] AND (((Data[6] OR ((Data[42] XOR ((Data[40] XOR Data[44]) XOR Data[19])) XOR Data[48])) XOR (((((NOT Data[35]) XOR ((Data[9] XOR Data[11]) XOR Data[20])) XOR ((Data[50] XOR Data[25]) XOR Data[1])) XOR (Data[6] OR ((Data[9] XOR Data[18]) XOR Data[18]))) XOR (((Data[44] AND Data[22]) XOR (NOT Data[9])) XOR Data[25]))) XOR (Data[26] AND Data[38]))))) OR (((TRUE AND (((((NOT (Data[23] OR Data[16])) AND (NOT ((Data[22] XOR Data[50]) XOR Data[9]))) XOR ((((NOT Data[42]) XOR (NOT Data[14])) XOR ((Data[3] XOR Data[34]) XOR Data[28])) OR (NOT (NOT Data[24])))) XOR ((Data[25] AND (Data[40] AND Data[13])) AND (Data[5] OR ((Data[10] XOR Data[1]) XOR Data[31])))) AND ((((NOT (Data[8] AND Data[33])) XOR (((Data[17] XOR Data[34]) XOR Data[34]) AND Data[6])) XOR (((Data[7] XOR Data[43]) XOR Data[13]) AND Data[11])) OR ((Data[34] XOR (NOT ((Data[41] XOR TRUE) XOR Data[49]))) XOR (((Data[39] XOR Data[49]) XOR Data[43]) AND ((Data[30] XOR Data[26]) XOR Data[36])))))) XOR (Data[41] AND (((((Data[18] OR FALSE) AND (Data[50] OR Data[45])) OR (((Data[9] OR Data[7]) XOR (NOT Data[18])) XOR (Data[34] OR Data[21]))) AND Data[6]) OR ((Data[40] XOR ((Data[7] XOR FALSE) XOR ((Data[17] AND Data[37]) AND Data[24]))) XOR ((NOT Data[16]) OR (NOT (Data[22] OR Data[8]))))))) XOR Data[16]))) XOR (Data[9] OR (NOT ((Data[8] XOR ((NOT ((((Data[18] OR Data[28]) XOR (Data[17] AND Data[6])) XOR (TRUE OR Data[4])) OR (NOT ((Data[26] XOR Data[22]) XOR Data[30])))) OR ((((NOT Data[4]) AND (((Data[48] OR Data[34]) XOR (Data[39] OR Data[15])) XOR (Data[41] AND Data[46]))) XOR (NOT (NOT (NOT Data[32])))) XOR (((NOT (NOT Data[13])) XOR Data[23]) XOR Data[8])))) XOR ((Data[9] XOR ((Data[35] AND (Data[3] AND (Data[43] OR Data[44]))) AND (Data[21] OR (Data[3] AND ((Data[4] XOR Data[50]) XOR Data[21]))))) XOR (((((Data[29] AND (NOT Data[40])) XOR (((Data[32] AND Data[21]) XOR (Data[10] AND Data[25])) XOR ((FALSE XOR Data[32]) XOR Data[24]))) XOR (NOT (Data[18] AND Data[45]))) XOR ((Data[46] AND (Data[27] AND Data[23])) OR Data[3])) XOR (((NOT (Data[32] OR Data[3])) XOR ((Data[48] AND Data[28]) OR (Data[18] AND Data[4]))) XOR (((Data[38] AND Data[23]) XOR (NOT Data[48])) XOR Data[1])))))))) OR (NOT ((((((Data[14] OR (((NOT (Data[18] AND Data[27])) XOR ((NOT Data[46]) OR (NOT Data[22]))) XOR ((NOT Data[15]) OR ((Data[27] XOR Data[25]) XOR Data[25])))) XOR ((((((((Data[48] XOR Data[20]) XOR Data[49]) XOR (NOT Data[6])) XOR (Data[21] OR Data[24])) XOR (NOT ((Data[45] XOR Data[13]) XOR Data[7]))) XOR (NOT Data[16])) XOR ((((Data[41] OR Data[27]) AND (Data[19] AND Data[19])) XOR Data[46]) XOR Data[49])) XOR (NOT Data[3]))) XOR Data[6]) OR (Data[18] AND (((((Data[35] AND Data[46]) OR (Data[19] OR Data[12])) XOR (NOT ((Data[35] XOR Data[22]) XOR Data[28]))) XOR ((Data[36] AND Data[18]) OR (NOT Data[43]))) AND (((((Data[40] XOR Data[26]) XOR Data[18]) XOR (Data[33] AND Data[31])) XOR (NOT Data[43])) AND (((Data[5] OR Data[20]) XOR Data[36]) XOR ((Data[18] XOR Data[49]) XOR Data[12])))))) OR Data[26]) AND Data[18])));
    OutReady := 1;
    CollectInput(RESET:=TRUE);
  END_IF;
END_PROGRAM

CONFIGURATION Config0
  RESOURCE Res0 ON PLC
    TASK task0(INTERVAL := T#20ms,PRIORITY := 0);
    PROGRAM instance0 WITH task0 : Boiler;
  END_RESOURCE
END_CONFIGURATION

(* ---- RND-EXPR_groan-hints-rogue.st ---- *)
(*
This code implements a randomly grown symbolic expression:

(!(false & IN38)) & (!(IN32))

*)

FUNCTION_BLOCK F_CollectInput
  VAR_IN_OUT
      Data : ARRAY[1..50] OF BOOL;
  END_VAR
  VAR_INPUT
      TICK  : BOOL := 0;
      IN1   : BOOL := 0;
      IN2   : BOOL := 0;
      IN3   : BOOL := 0;
      IN4   : BOOL := 0;
      IN5   : BOOL := 0;
      RESET : BOOL := FALSE;
  END_VAR
  VAR_OUTPUT
      Finished : BOOL;
  END_VAR
  VAR
      j    : USINT := 1;
      tock : BOOL  := 0;
  END_VAR
  IF NOT RESET AND tock = NOT TICK THEN
      Data[j]   := IN1;
      Data[j+1] := IN2;
      Data[j+2] := IN3;
      Data[j+3] := IN4;
      Data[j+4] := IN5;
      j := j + 5;
      tock := TICK;
  ELSE
      j := 1;
      tock := 0;
  END_IF;
  Finished := (j > 50);
END_FUNCTION_BLOCK

PROGRAM Boiler
  VAR
    Data  : ARRAY[1..50] OF BOOL;
    Ready : BOOL;
    CollectInput : F_CollectInput;
  END_VAR
  VAR
    TICK     AT %IX1.0 : BOOL;
    IN1      AT %IX0.3 : BOOL;
    IN2      AT %IX0.4 : BOOL;
    IN3      AT %IX0.5 : BOOL;
    IN4      AT %IX0.6 : BOOL;
    IN5      AT %IX0.7 : BOOL;
    OutReady AT %QX0.0 : BOOL := FALSE;
    FeedNext AT %QX0.1 : BOOL := FALSE;
    Out      AT %QX0.2 : BOOL;
  END_VAR
  CollectInput(TICK:=TICK, IN1:=IN1, IN2:=IN2, IN3:=IN3, IN4:=IN4, IN5:=IN5);
  Ready := CollectInput.Finished;
  FeedNext := 1;
  IF Ready THEN
    Out := ((NOT (FALSE AND Data[38])) AND (NOT Data[32]));
    OutReady := 1;
    CollectInput(RESET:=TRUE);
  END_IF;
END_PROGRAM

CONFIGURATION Config0
  RESOURCE Res0 ON PLC
    TASK task0(INTERVAL := T#20ms,PRIORITY := 0);
    PROGRAM instance0 WITH task0 : Boiler;
  END_RESOURCE
END_CONFIGURATION

(* ---- RND-EXPR_guilt-fames-dined.st ---- *)
(*
This code implements a randomly grown symbolic expression:

((((!(xor(xor(!(!((IN22 | IN39) | (IN19 | IN48))), IN37 & (!(IN40))), !(IN3 & IN44)))) | (!(xor(xor(xor(xor(xor(xor((!(IN22)) | (IN11 & IN37), true), IN25), xor(xor(xor(xor(IN7 | IN32, IN16 & IN30), IN31 | IN37), IN43 & (IN9 & IN6)), (xor(xor(IN27, IN23), IN5)) | (IN20 | IN42))), (IN13 | IN11) & (xor(xor(IN11 | IN34, IN4 & IN43), xor(xor(IN12, IN48), IN41)))), xor(xor(((!(IN7)) & IN8) | ((xor(xor(IN12, IN26), IN15)) | IN41), (!(IN22 & IN47)) & (!(IN28 | IN40))), (xor(xor(IN22, IN22 | IN41), IN4)) | ((xor(xor(IN24, IN45), IN6)) & (IN23 & IN38)))), xor(xor(!(!(xor(xor(IN2, IN39), IN43))), IN13), !((xor(true, IN6)) & (!(IN4)))))))) | ((xor(xor(xor(xor((xor(xor(IN8, !(IN50)), (!(IN34)) & (!(IN32)))) | ((IN2 | (IN8 | IN46)) & (!(IN12 | IN41))), IN6 | IN26), !(((IN30 & IN2) | IN20) | IN32)), IN29), ((IN15 | ((IN38 | IN21) & (!(IN6)))) & IN35) | ((!((!(IN28)) & (IN33 | IN20))) | (xor(xor(xor(xor(xor(xor(IN27, IN30), IN43), xor(xor(IN12, IN23), IN31)), xor(xor(IN1, IN44), IN33)), !(!(IN2))), xor(xor(IN9 & IN13, xor(xor(IN2, IN49), IN11)), IN18 & IN28)))))) | (((!(xor(xor(xor(xor(IN11 | IN12, !(IN5)), IN9 & IN5), !(xor(xor(IN2, IN37), IN47))), xor(xor(!(IN34), IN31 & IN34), xor(xor(IN45, IN43), IN49))))) & (IN34 & (xor(xor(IN15, IN26), IN10 & (xor(xor(IN17, IN8), IN40)))))) | ((((xor(xor(!(IN38), !(IN33)), IN2)) & ((xor(xor(IN31, IN36), IN34)) | (IN13 | IN21))) | (IN26 | IN27)) | (!(IN32)))))) | (!((((xor(xor(xor(xor((!(IN33)) | (!(IN4)), IN25 | IN39), (!(IN31)) & (!(IN21))), ((IN20 & IN12) & (xor(xor(IN34, IN14), IN18))) & ((xor(false, IN11)) & IN22)), !(!(IN31)))) & (IN17 | (((IN20 & IN21) & (IN33 & IN15)) | IN10))) & (!(IN32))) | IN39))) | (!(xor(xor((true | IN39) & (xor(xor(xor(xor(xor(xor((xor(xor(!(IN30), IN36), IN7 | IN28)) | IN31, IN13), xor(xor(IN33 & (xor(xor(IN50, IN11), IN43)), !(!(IN35))), (xor(xor(IN30, false), IN35)) | IN10)), xor(xor((!(IN21 | IN50)) | ((xor(xor(IN6, IN9), IN9)) | (!(IN44))), (xor(xor(IN2 & IN22, IN4 | IN20), xor(xor(IN21, IN32), false))) & (!(!(IN26)))), xor(xor(xor(xor(IN16 & IN21, IN48), IN34 | IN3), !(xor(xor(IN19, IN19), IN44))), !(xor(xor(IN25, IN29), IN4))))), IN46 & ((!(IN3 & IN29)) | IN38)), (xor(xor((IN33 & (xor(xor(IN38, IN14), IN22))) | ((xor(xor(IN38, IN23), IN46)) | (xor(xor(IN37, IN32), IN24))), xor(xor(IN31 & (IN5 | IN29), xor(xor(IN12, xor(xor(false, IN36), IN10)), !(IN37))), xor(xor(IN50 | IN45, xor(xor(IN34, IN17), IN17)), IN5))), !(xor(xor(IN34 | IN16, xor(xor(IN48, IN30), IN43)), IN36 | IN29)))) & IN11), ((!((xor(xor(IN32, IN13), IN39)) & (xor(xor(IN42, IN16), IN20)))) | (IN22 & (xor(xor(IN1 | IN3, xor(xor(IN43, true), IN45)), IN4 & IN29)))) & (xor(xor(xor(xor(IN12 | (IN45 | IN48), xor(xor(!(IN32), true), xor(xor(IN7, IN20), IN47))), xor(xor(IN40 | IN29, IN22 | IN32), xor(xor(IN21, IN16), true))), IN30), IN42)))), xor(xor((xor(xor(xor(xor(((xor(xor(IN1, IN30), IN45)) & IN38) | (xor(xor(IN19 & IN48, xor(xor(IN26, IN2), IN10)), IN36 & IN24)), xor(xor((IN15 | true) | (!(IN17)), IN30), IN18 | (xor(xor(IN48, IN31), IN28)))), (xor(xor(xor(xor(IN47, false), IN32), IN37 | IN28), IN15 | IN26)) & IN15), IN15), IN45 | (!(IN49)))) | (IN39 & ((xor(xor(!(IN21), xor(xor(IN24 | IN30, IN11 | IN22), IN20)), (IN36 & IN28) & (xor(xor(IN44, IN7), IN37)))) & (xor(xor((!(IN24)) & (!(IN38)), (IN47 | IN12) & (IN28 & IN16)), (false | IN24) | IN33)))), IN19), IN39 & IN8)), !(!(xor(xor(xor(xor(xor(xor(!(IN29), !(xor(xor(IN26, IN31), IN44))), (!(IN32)) | (IN5 | IN8)), (xor(xor(!(IN8), IN14), IN17 & IN31)) | (!(IN25 & IN1))), IN11), (xor(xor(xor(xor(IN29 | IN47, IN36 | IN27), IN13), IN41), xor(xor(IN23 & IN50, xor(xor(IN18, IN27), IN28)), IN11 | IN11))) | (!((IN36 | IN47) | IN23))), !(xor(xor((IN17 & IN18) & (!(IN21)), xor(xor(IN5 | false, IN15 | IN48), IN47 | IN22)), xor(xor(IN1, false | IN8), xor(xor(IN36, IN33), IN31))))))))))

*)

FUNCTION_BLOCK F_CollectInput
  VAR_IN_OUT
      Data : ARRAY[1..50] OF BOOL;
  END_VAR
  VAR_INPUT
      TICK  : BOOL := 0;
      IN1   : BOOL := 0;
      IN2   : BOOL := 0;
      IN3   : BOOL := 0;
      IN4   : BOOL := 0;
      IN5   : BOOL := 0;
      RESET : BOOL := FALSE;
  END_VAR
  VAR_OUTPUT
      Finished : BOOL;
  END_VAR
  VAR
      j    : USINT := 1;
      tock : BOOL  := 0;
  END_VAR
  IF NOT RESET AND tock = NOT TICK THEN
      Data[j]   := IN1;
      Data[j+1] := IN2;
      Data[j+2] := IN3;
      Data[j+3] := IN4;
      Data[j+4] := IN5;
      j := j + 5;
      tock := TICK;
  ELSE
      j := 1;
      tock := 0;
  END_IF;
  Finished := (j > 50);
END_FUNCTION_BLOCK

PROGRAM Boiler
  VAR
    Data  : ARRAY[1..50] OF BOOL;
    Ready : BOOL;
    CollectInput : F_CollectInput;
  END_VAR
  VAR
    TICK     AT %IX1.0 : BOOL;
    IN1      AT %IX0.3 : BOOL;
    IN2      AT %IX0.4 : BOOL;
    IN3      AT %IX0.5 : BOOL;
    IN4      AT %IX0.6 : BOOL;
    IN5      AT %IX0.7 : BOOL;
    OutReady AT %QX0.0 : BOOL := FALSE;
    FeedNext AT %QX0.1 : BOOL := FALSE;
    Out      AT %QX0.2 : BOOL;
  END_VAR
  CollectInput(TICK:=TICK, IN1:=IN1, IN2:=IN2, IN3:=IN3, IN4:=IN4, IN5:=IN5);
  Ready := CollectInput.Finished;
  FeedNext := 1;
  IF Ready THEN
    Out := (((((NOT (((NOT (NOT ((Data[22] OR Data[39]) OR (Data[19] OR Data[48])))) XOR (Data[37] AND (NOT Data[40]))) XOR (NOT (Data[3] AND Data[44])))) OR (NOT ((((((((NOT Data[22]) OR (Data[11] AND Data[37])) XOR TRUE) XOR Data[25]) XOR (((((Data[7] OR Data[32]) XOR (Data[16] AND Data[30])) XOR (Data[31] OR Data[37])) XOR (Data[43] AND (Data[9] AND Data[6]))) XOR (((Data[27] XOR Data[23]) XOR Data[5]) OR (Data[20] OR Data[42])))) XOR ((Data[13] OR Data[11]) AND (((Data[11] OR Data[34]) XOR (Data[4] AND Data[43])) XOR ((Data[12] XOR Data[48]) XOR Data[41])))) XOR (((((NOT Data[7]) AND Data[8]) OR (((Data[12] XOR Data[26]) XOR Data[15]) OR Data[41])) XOR ((NOT (Data[22] AND Data[47])) AND (NOT (Data[28] OR Data[40])))) XOR (((Data[22] XOR (Data[22] OR Data[41])) XOR Data[4]) OR (((Data[24] XOR Data[45]) XOR Data[6]) AND (Data[23] AND Data[38]))))) XOR (((NOT (NOT ((Data[2] XOR Data[39]) XOR Data[43]))) XOR Data[13]) XOR (NOT ((TRUE XOR Data[6]) AND (NOT Data[4]))))))) OR ((((((((Data[8] XOR (NOT Data[50])) XOR ((NOT Data[34]) AND (NOT Data[32]))) OR ((Data[2] OR (Data[8] OR Data[46])) AND (NOT (Data[12] OR Data[41])))) XOR (Data[6] OR Data[26])) XOR (NOT (((Data[30] AND Data[2]) OR Data[20]) OR Data[32]))) XOR Data[29]) XOR (((Data[15] OR ((Data[38] OR Data[21]) AND (NOT Data[6]))) AND Data[35]) OR ((NOT ((NOT Data[28]) AND (Data[33] OR Data[20]))) OR ((((((Data[27] XOR Data[30]) XOR Data[43]) XOR ((Data[12] XOR Data[23]) XOR Data[31])) XOR ((Data[1] XOR Data[44]) XOR Data[33])) XOR (NOT (NOT Data[2]))) XOR (((Data[9] AND Data[13]) XOR ((Data[2] XOR Data[49]) XOR Data[11])) XOR (Data[18] AND Data[28])))))) OR (((NOT (((((Data[11] OR Data[12]) XOR (NOT Data[5])) XOR (Data[9] AND Data[5])) XOR (NOT ((Data[2] XOR Data[37]) XOR Data[47]))) XOR (((NOT Data[34]) XOR (Data[31] AND Data[34])) XOR ((Data[45] XOR Data[43]) XOR Data[49])))) AND (Data[34] AND ((Data[15] XOR Data[26]) XOR (Data[10] AND ((Data[17] XOR Data[8]) XOR Data[40]))))) OR ((((((NOT Data[38]) XOR (NOT Data[33])) XOR Data[2]) AND (((Data[31] XOR Data[36]) XOR Data[34]) OR (Data[13] OR Data[21]))) OR (Data[26] OR Data[27])) OR (NOT Data[32]))))) OR (NOT (((((((((NOT Data[33]) OR (NOT Data[4])) XOR (Data[25] OR Data[39])) XOR ((NOT Data[31]) AND (NOT Data[21]))) XOR (((Data[20] AND Data[12]) AND ((Data[34] XOR Data[14]) XOR Data[18])) AND ((FALSE XOR Data[11]) AND Data[22]))) XOR (NOT (NOT Data[31]))) AND (Data[17] OR (((Data[20] AND Data[21]) AND (Data[33] AND Data[15])) OR Data[10]))) AND (NOT Data[32])) OR Data[39]))) OR (NOT ((((TRUE OR Data[39]) AND ((((((((((NOT Data[30]) XOR Data[36]) XOR (Data[7] OR Data[28])) OR Data[31]) XOR Data[13]) XOR (((Data[33] AND ((Data[50] XOR Data[11]) XOR Data[43])) XOR (NOT (NOT Data[35]))) XOR (((Data[30] XOR FALSE) XOR Data[35]) OR Data[10]))) XOR ((((NOT (Data[21] OR Data[50])) OR (((Data[6] XOR Data[9]) XOR Data[9]) OR (NOT Data[44]))) XOR ((((Data[2] AND Data[22]) XOR (Data[4] OR Data[20])) XOR ((Data[21] XOR Data[32]) XOR FALSE)) AND (NOT (NOT Data[26])))) XOR (((((Data[16] AND Data[21]) XOR Data[48]) XOR (Data[34] OR Data[3])) XOR (NOT ((Data[19] XOR Data[19]) XOR Data[44]))) XOR (NOT ((Data[25] XOR Data[29]) XOR Data[4]))))) XOR (Data[46] AND ((NOT (Data[3] AND Data[29])) OR Data[38]))) XOR (((((Data[33] AND ((Data[38] XOR Data[14]) XOR Data[22])) OR (((Data[38] XOR Data[23]) XOR Data[46]) OR ((Data[37] XOR Data[32]) XOR Data[24]))) XOR (((Data[31] AND (Data[5] OR Data[29])) XOR ((Data[12] XOR ((FALSE XOR Data[36]) XOR Data[10])) XOR (NOT Data[37]))) XOR (((Data[50] OR Data[45]) XOR ((Data[34] XOR Data[17]) XOR Data[17])) XOR Data[5]))) XOR (NOT (((Data[34] OR Data[16]) XOR ((Data[48] XOR Data[30]) XOR Data[43])) XOR (Data[36] OR Data[29])))) AND Data[11])) XOR (((NOT (((Data[32] XOR Data[13]) XOR Data[39]) AND ((Data[42] XOR Data[16]) XOR Data[20]))) OR (Data[22] AND (((Data[1] OR Data[3]) XOR ((Data[43] XOR TRUE) XOR Data[45])) XOR (Data[4] AND Data[29])))) AND (((((Data[12] OR (Data[45] OR Data[48])) XOR (((NOT Data[32]) XOR TRUE) XOR ((Data[7] XOR Data[20]) XOR Data[47]))) XOR (((Data[40] OR Data[29]) XOR (Data[22] OR Data[32])) XOR ((Data[21] XOR Data[16]) XOR TRUE))) XOR Data[30]) XOR Data[42])))) XOR (((((((((((Data[1] XOR Data[30]) XOR Data[45]) AND Data[38]) OR (((Data[19] AND Data[48]) XOR ((Data[26] XOR Data[2]) XOR Data[10])) XOR (Data[36] AND Data[24]))) XOR ((((Data[15] OR TRUE) OR (NOT Data[17])) XOR Data[30]) XOR (Data[18] OR ((Data[48] XOR Data[31]) XOR Data[28])))) XOR (((((Data[47] XOR FALSE) XOR Data[32]) XOR (Data[37] OR Data[28])) XOR (Data[15] OR Data[26])) AND Data[15])) XOR Data[15]) XOR (Data[45] OR (NOT Data[49]))) OR (Data[39] AND ((((NOT Data[21]) XOR (((Data[24] OR Data[30]) XOR (Data[11] OR Data[22])) XOR Data[20])) XOR ((Data[36] AND Data[28]) AND ((Data[44] XOR Data[7]) XOR Data[37]))) AND ((((NOT Data[24]) AND (NOT Data[38])) XOR ((Data[47] OR Data[12]) AND (Data[28] AND Data[16]))) XOR ((FALSE OR Data[24]) OR Data[33]))))) XOR Data[19]) XOR (Data[39] AND Data[8]))) XOR (NOT (NOT (((((((NOT Data[29]) XOR (NOT ((Data[26] XOR Data[31]) XOR Data[44]))) XOR ((NOT Data[32]) OR (Data[5] OR Data[8]))) XOR ((((NOT Data[8]) XOR Data[14]) XOR (Data[17] AND Data[31])) OR (NOT (Data[25] AND Data[1])))) XOR Data[11]) XOR ((((((Data[29] OR Data[47]) XOR (Data[36] OR Data[27])) XOR Data[13]) XOR Data[41]) XOR (((Data[23] AND Data[50]) XOR ((Data[18] XOR Data[27]) XOR Data[28])) XOR (Data[11] OR Data[11]))) OR (NOT ((Data[36] OR Data[47]) OR Data[23])))) XOR (NOT ((((Data[17] AND Data[18]) AND (NOT Data[21])) XOR (((Data[5] OR FALSE) XOR (Data[15] OR Data[48])) XOR (Data[47] OR Data[22]))) XOR ((Data[1] XOR (FALSE OR Data[8])) XOR ((Data[36] XOR Data[33]) XOR Data[31]))))))))));
    OutReady := 1;
    CollectInput(RESET:=TRUE);
  END_IF;
END_PROGRAM

CONFIGURATION Config0
  RESOURCE Res0 ON PLC
    TASK task0(INTERVAL := T#20ms,PRIORITY := 0);
    PROGRAM instance0 WITH task0 : Boiler;
  END_RESOURCE
END_CONFIGURATION

(* ---- RND-EXPR_happy-patio-shuck.st ---- *)
(*
This code implements a randomly grown symbolic expression:

xor(xor((xor(xor((!(xor(xor(IN1, !(((xor(xor(IN9, false), IN23)) | (!(IN25))) & IN44)), (!(IN16 | (IN48 | IN3))) & ((!(IN24)) | ((IN45 | IN50) & (xor(xor(true, IN37), IN36))))))) | (!(xor(xor(IN45, !(!(IN24 | (xor(xor(IN42, IN24), IN37))))), xor(xor(IN32 | (xor(xor(!(IN31), IN1 | IN43), IN50 & IN38)), ((!(IN37)) | (IN24 | IN12)) & (xor(xor(xor(xor(IN23, IN20), IN44), IN3 & IN28), xor(xor(IN4, IN33), IN46)))), !((IN44 & IN24) & (!(IN26))))))), IN48), !(xor(xor(IN19, IN41), IN10 & (xor(xor(!((IN31 | IN33) | (!(IN2))), IN49), ((IN33 & IN10) & (!(IN46))) & (xor(xor(IN48, !(IN17)), IN17 | IN23)))))))) | IN35, (!((xor(xor(xor(xor(!(((!(IN13)) | (IN33 & IN11)) | ((!(IN26)) & (IN31 & IN33))), ((IN13 | (IN37 & IN1)) & (IN15 & (xor(xor(IN18, IN36), IN22)))) | (!(IN32 | (IN20 | IN32)))), (((xor(xor(IN43, IN21), false)) | IN15) | ((xor(xor(IN8, IN50), IN26)) | (xor(xor(IN42, IN47), IN44)))) | ((!(xor(xor(IN45, IN2), IN34))) | ((!(IN9)) | (!(IN18))))), !(xor(xor(!((xor(xor(IN42, IN48), IN14)) & (IN12 | IN49)), IN38), IN46))), xor(xor(xor(xor(IN23, (!(IN16)) & ((IN30 & IN49) | (xor(xor(IN44, IN3), IN22)))), !(!(xor(xor(IN5, IN31), IN5)))), IN13 | (!((!(IN7)) | IN1))), ((xor(xor(IN2 | IN24, IN44 & IN38), IN46 | IN31)) | ((IN6 & IN11) | IN18)) | ((xor(xor(!(IN49), xor(xor(IN4, IN36), IN32)), xor(xor(IN18, IN24), IN30))) | ((IN19 | IN34) | (xor(xor(IN35, IN12), IN45))))))) & IN21)) & ((xor(xor((IN19 | IN26) & IN27, (xor(xor(xor(xor(IN7 | ((!(IN50)) | (xor(xor(IN9, IN33), IN2))), !(!(xor(xor(IN14, IN12), IN17)))), IN31), (!((!(IN39)) | (xor(xor(IN24, IN35), IN23)))) | (xor(xor((IN18 & IN8) & (xor(xor(IN46, IN25), IN35)), (IN17 & IN41) & false), xor(xor(!(IN15), xor(xor(IN34, IN35), IN1)), IN27 | IN35)))), xor(xor((xor(xor(xor(xor(IN24, IN41), IN40), IN5 | IN46), !(IN10))) & ((xor(xor(IN32, IN9), IN10)) | (IN32 & false)), xor(xor(xor(xor(!(IN32), IN15 | IN40), IN7 & IN30), (IN37 & IN11) & (IN19 | IN42)), !(!(IN46)))), IN2))) | ((!(!(!(IN23 & IN25)))) & IN39)), IN2)) | IN19)), !(!(IN5 & IN24)))

*)

FUNCTION_BLOCK F_CollectInput
  VAR_IN_OUT
      Data : ARRAY[1..50] OF BOOL;
  END_VAR
  VAR_INPUT
      TICK  : BOOL := 0;
      IN1   : BOOL := 0;
      IN2   : BOOL := 0;
      IN3   : BOOL := 0;
      IN4   : BOOL := 0;
      IN5   : BOOL := 0;
      RESET : BOOL := FALSE;
  END_VAR
  VAR_OUTPUT
      Finished : BOOL;
  END_VAR
  VAR
      j    : USINT := 1;
      tock : BOOL  := 0;
  END_VAR
  IF NOT RESET AND tock = NOT TICK THEN
      Data[j]   := IN1;
      Data[j+1] := IN2;
      Data[j+2] := IN3;
      Data[j+3] := IN4;
      Data[j+4] := IN5;
      j := j + 5;
      tock := TICK;
  ELSE
      j := 1;
      tock := 0;
  END_IF;
  Finished := (j > 50);
END_FUNCTION_BLOCK

PROGRAM Boiler
  VAR
    Data  : ARRAY[1..50] OF BOOL;
    Ready : BOOL;
    CollectInput : F_CollectInput;
  END_VAR
  VAR
    TICK     AT %IX1.0 : BOOL;
    IN1      AT %IX0.3 : BOOL;
    IN2      AT %IX0.4 : BOOL;
    IN3      AT %IX0.5 : BOOL;
    IN4      AT %IX0.6 : BOOL;
    IN5      AT %IX0.7 : BOOL;
    OutReady AT %QX0.0 : BOOL := FALSE;
    FeedNext AT %QX0.1 : BOOL := FALSE;
    Out      AT %QX0.2 : BOOL;
  END_VAR
  CollectInput(TICK:=TICK, IN1:=IN1, IN2:=IN2, IN3:=IN3, IN4:=IN4, IN5:=IN5);
  Ready := CollectInput.Finished;
  FeedNext := 1;
  IF Ready THEN
    Out := (((((((NOT ((Data[1] XOR (NOT ((((Data[9] XOR FALSE) XOR Data[23]) OR (NOT Data[25])) AND Data[44]))) XOR ((NOT (Data[16] OR (Data[48] OR Data[3]))) AND ((NOT Data[24]) OR ((Data[45] OR Data[50]) AND ((TRUE XOR Data[37]) XOR Data[36])))))) OR (NOT ((Data[45] XOR (NOT (NOT (Data[24] OR ((Data[42] XOR Data[24]) XOR Data[37]))))) XOR (((Data[32] OR (((NOT Data[31]) XOR (Data[1] OR Data[43])) XOR (Data[50] AND Data[38]))) XOR (((NOT Data[37]) OR (Data[24] OR Data[12])) AND ((((Data[23] XOR Data[20]) XOR Data[44]) XOR (Data[3] AND Data[28])) XOR ((Data[4] XOR Data[33]) XOR Data[46])))) XOR (NOT ((Data[44] AND Data[24]) AND (NOT Data[26]))))))) XOR Data[48]) XOR (NOT ((Data[19] XOR Data[41]) XOR (Data[10] AND (((NOT ((Data[31] OR Data[33]) OR (NOT Data[2]))) XOR Data[49]) XOR (((Data[33] AND Data[10]) AND (NOT Data[46])) AND ((Data[48] XOR (NOT Data[17])) XOR (Data[17] OR Data[23])))))))) OR Data[35]) XOR ((NOT ((((((NOT (((NOT Data[13]) OR (Data[33] AND Data[11])) OR ((NOT Data[26]) AND (Data[31] AND Data[33])))) XOR (((Data[13] OR (Data[37] AND Data[1])) AND (Data[15] AND ((Data[18] XOR Data[36]) XOR Data[22]))) OR (NOT (Data[32] OR (Data[20] OR Data[32]))))) XOR (((((Data[43] XOR Data[21]) XOR FALSE) OR Data[15]) OR (((Data[8] XOR Data[50]) XOR Data[26]) OR ((Data[42] XOR Data[47]) XOR Data[44]))) OR ((NOT ((Data[45] XOR Data[2]) XOR Data[34])) OR ((NOT Data[9]) OR (NOT Data[18]))))) XOR (NOT (((NOT (((Data[42] XOR Data[48]) XOR Data[14]) AND (Data[12] OR Data[49]))) XOR Data[38]) XOR Data[46]))) XOR ((((Data[23] XOR ((NOT Data[16]) AND ((Data[30] AND Data[49]) OR ((Data[44] XOR Data[3]) XOR Data[22])))) XOR (NOT (NOT ((Data[5] XOR Data[31]) XOR Data[5])))) XOR (Data[13] OR (NOT ((NOT Data[7]) OR Data[1])))) XOR (((((Data[2] OR Data[24]) XOR (Data[44] AND Data[38])) XOR (Data[46] OR Data[31])) OR ((Data[6] AND Data[11]) OR Data[18])) OR ((((NOT Data[49]) XOR ((Data[4] XOR Data[36]) XOR Data[32])) XOR ((Data[18] XOR Data[24]) XOR Data[30])) OR ((Data[19] OR Data[34]) OR ((Data[35] XOR Data[12]) XOR Data[45])))))) AND Data[21])) AND (((((Data[19] OR Data[26]) AND Data[27]) XOR ((((((Data[7] OR ((NOT Data[50]) OR ((Data[9] XOR Data[33]) XOR Data[2]))) XOR (NOT (NOT ((Data[14] XOR Data[12]) XOR Data[17])))) XOR Data[31]) XOR ((NOT ((NOT Data[39]) OR ((Data[24] XOR Data[35]) XOR Data[23]))) OR ((((Data[18] AND Data[8]) AND ((Data[46] XOR Data[25]) XOR Data[35])) XOR ((Data[17] AND Data[41]) AND FALSE)) XOR (((NOT Data[15]) XOR ((Data[34] XOR Data[35]) XOR Data[1])) XOR (Data[27] OR Data[35]))))) XOR (((((((Data[24] XOR Data[41]) XOR Data[40]) XOR (Data[5] OR Data[46])) XOR (NOT Data[10])) AND (((Data[32] XOR Data[9]) XOR Data[10]) OR (Data[32] AND FALSE))) XOR (((((NOT Data[32]) XOR (Data[15] OR Data[40])) XOR (Data[7] AND Data[30])) XOR ((Data[37] AND Data[11]) AND (Data[19] OR Data[42]))) XOR (NOT (NOT Data[46])))) XOR Data[2])) OR ((NOT (NOT (NOT (Data[23] AND Data[25])))) AND Data[39]))) XOR Data[2]) OR Data[19]))) XOR (NOT (NOT (Data[5] AND Data[24]))));
    OutReady := 1;
    CollectInput(RESET:=TRUE);
  END_IF;
END_PROGRAM

CONFIGURATION Config0
  RESOURCE Res0 ON PLC
    TASK task0(INTERVAL := T#20ms,PRIORITY := 0);
    PROGRAM instance0 WITH task0 : Boiler;
  END_RESOURCE
END_CONFIGURATION

(* ---- RND-EXPR_helps-sound-boast.st ---- *)
(*
This code implements a randomly grown symbolic expression:

!(xor(xor((xor(xor((IN49 | (xor(xor(!(xor(xor(xor(xor(IN8, IN35), IN20), xor(xor(IN46, IN3), IN36)), !(IN18))), !(IN46)), !(xor(xor(IN45, !(IN41)), IN31 & IN32))))) | ((IN26 & IN5) | ((!((!(IN32)) | (IN35 & IN13))) | (!(!(!(IN14)))))), (!(xor(xor(IN3, IN23), IN36 & (IN21 | IN45)))) | IN1), ((xor(xor(IN5, IN47 & ((!(IN48)) | (IN29 | IN37))), !(IN20))) & (!((xor(xor(IN39 | IN3, IN18 & IN8), !(IN47))) | (IN5 & (xor(xor(IN42, IN8), IN34)))))) | ((!((!(!(IN31))) | ((xor(xor(IN42, IN50), IN50)) & (IN15 & IN15)))) & ((!((IN48 & IN15) & IN8)) & (xor(xor((xor(xor(IN21, IN23), IN32)) | IN33, xor(xor(IN2 & IN1, xor(xor(IN45, IN16), IN27)), IN2 & IN16)), xor(xor(IN50, IN8), !(IN6)))))))) | (!(IN5 | ((xor(xor((IN40 | IN10) | IN42, !(xor(xor(!(IN24), IN2 & IN21), IN41 | IN36))), !(IN19))) | (IN30 | (xor(xor((IN47 & IN33) | (!(IN15)), (!(IN47)) & (IN25 | IN8)), (IN42 & IN6) | (IN37 & IN25))))))), xor(xor(xor(xor(xor(xor((IN5 | ((IN44 & (IN1 & IN11)) & (!(IN26 | IN47)))) & (((!(xor(xor(IN16, IN7), IN43))) | (!(xor(xor(false, IN28), IN46)))) & (xor(xor(!(xor(xor(IN21, IN34), IN39)), !(IN26 | IN34)), (IN1 & IN44) & (xor(xor(IN43, IN1), IN47))))), ((!(!(IN32))) | (!(IN5 & IN31))) & (!(xor(xor((xor(xor(IN30, IN30), IN37)) & (IN13 & IN50), IN42), (xor(xor(IN20, IN44), IN30)) | (IN13 | IN32))))), IN26), (IN16 | ((IN18 & ((IN38 & IN9) & (xor(xor(IN34, IN26), IN40)))) & ((!(IN18)) & ((xor(xor(IN45, true), IN2)) | (!(IN16)))))) | IN35), IN30), ((!(!(xor(xor(xor(xor(IN13 & IN10, xor(xor(false, IN33), IN21)), !(IN8)), xor(xor(!(IN35), IN35), IN33 | IN9)), !(!(IN34)))))) | IN29) | (!(IN21 | ((((xor(xor(IN25, IN33), IN4)) & (!(IN26))) & (!(IN11))) & ((xor(xor(IN43, !(IN3)), false)) | (!(IN22 | IN8))))))), !(IN41))), ((!(((!(xor(xor(IN15 & true, IN6), IN48 & IN46))) | (!(IN44 & (IN19 & IN30)))) & ((!(xor(xor(IN45 & IN3, IN28), IN47 & IN44))) & IN20))) | IN46) | ((xor(xor(IN27, xor(xor(!((IN10 | IN27) | (IN24 | (IN38 | IN33))), IN37 & (IN7 | (xor(xor(!(IN46), xor(xor(IN20, IN42), IN46)), IN10)))), IN15 & (xor(xor((xor(xor(false, IN15), IN41)) | (IN19 & IN28), IN25 | (IN48 | IN14)), !(!(IN38)))))), IN9)) & (xor(xor((!((xor(xor(IN2 | IN41, IN15 & IN50), IN39 | IN34)) | ((xor(xor(IN50, IN15), IN2)) | (!(IN36))))) & IN11, !((!(IN26 & (IN10 & IN45))) & (!(IN19)))), (IN13 & (IN45 | (xor(xor(IN42 | IN30, IN44 & true), !(IN46))))) | (IN19 & ((!(xor(xor(IN26, IN9), IN43))) & ((!(IN29)) | (xor(xor(IN11, IN23), false))))))))))

*)

FUNCTION_BLOCK F_CollectInput
  VAR_IN_OUT
      Data : ARRAY[1..50] OF BOOL;
  END_VAR
  VAR_INPUT
      TICK  : BOOL := 0;
      IN1   : BOOL := 0;
      IN2   : BOOL := 0;
      IN3   : BOOL := 0;
      IN4   : BOOL := 0;
      IN5   : BOOL := 0;
      RESET : BOOL := FALSE;
  END_VAR
  VAR_OUTPUT
      Finished : BOOL;
  END_VAR
  VAR
      j    : USINT := 1;
      tock : BOOL  := 0;
  END_VAR
  IF NOT RESET AND tock = NOT TICK THEN
      Data[j]   := IN1;
      Data[j+1] := IN2;
      Data[j+2] := IN3;
      Data[j+3] := IN4;
      Data[j+4] := IN5;
      j := j + 5;
      tock := TICK;
  ELSE
      j := 1;
      tock := 0;
  END_IF;
  Finished := (j > 50);
END_FUNCTION_BLOCK

PROGRAM Boiler
  VAR
    Data  : ARRAY[1..50] OF BOOL;
    Ready : BOOL;
    CollectInput : F_CollectInput;
  END_VAR
  VAR
    TICK     AT %IX1.0 : BOOL;
    IN1      AT %IX0.3 : BOOL;
    IN2      AT %IX0.4 : BOOL;
    IN3      AT %IX0.5 : BOOL;
    IN4      AT %IX0.6 : BOOL;
    IN5      AT %IX0.7 : BOOL;
    OutReady AT %QX0.0 : BOOL := FALSE;
    FeedNext AT %QX0.1 : BOOL := FALSE;
    Out      AT %QX0.2 : BOOL;
  END_VAR
  CollectInput(TICK:=TICK, IN1:=IN1, IN2:=IN2, IN3:=IN3, IN4:=IN4, IN5:=IN5);
  Ready := CollectInput.Finished;
  FeedNext := 1;
  IF Ready THEN
    Out := (NOT (((((((Data[49] OR (((NOT ((((Data[8] XOR Data[35]) XOR Data[20]) XOR ((Data[46] XOR Data[3]) XOR Data[36])) XOR (NOT Data[18]))) XOR (NOT Data[46])) XOR (NOT ((Data[45] XOR (NOT Data[41])) XOR (Data[31] AND Data[32]))))) OR ((Data[26] AND Data[5]) OR ((NOT ((NOT Data[32]) OR (Data[35] AND Data[13]))) OR (NOT (NOT (NOT Data[14])))))) XOR ((NOT ((Data[3] XOR Data[23]) XOR (Data[36] AND (Data[21] OR Data[45])))) OR Data[1])) XOR ((((Data[5] XOR (Data[47] AND ((NOT Data[48]) OR (Data[29] OR Data[37])))) XOR (NOT Data[20])) AND (NOT ((((Data[39] OR Data[3]) XOR (Data[18] AND Data[8])) XOR (NOT Data[47])) OR (Data[5] AND ((Data[42] XOR Data[8]) XOR Data[34]))))) OR ((NOT ((NOT (NOT Data[31])) OR (((Data[42] XOR Data[50]) XOR Data[50]) AND (Data[15] AND Data[15])))) AND ((NOT ((Data[48] AND Data[15]) AND Data[8])) AND (((((Data[21] XOR Data[23]) XOR Data[32]) OR Data[33]) XOR (((Data[2] AND Data[1]) XOR ((Data[45] XOR Data[16]) XOR Data[27])) XOR (Data[2] AND Data[16]))) XOR ((Data[50] XOR Data[8]) XOR (NOT Data[6]))))))) OR (NOT (Data[5] OR (((((Data[40] OR Data[10]) OR Data[42]) XOR (NOT (((NOT Data[24]) XOR (Data[2] AND Data[21])) XOR (Data[41] OR Data[36])))) XOR (NOT Data[19])) OR (Data[30] OR ((((Data[47] AND Data[33]) OR (NOT Data[15])) XOR ((NOT Data[47]) AND (Data[25] OR Data[8]))) XOR ((Data[42] AND Data[6]) OR (Data[37] AND Data[25])))))))) XOR ((((((((Data[5] OR ((Data[44] AND (Data[1] AND Data[11])) AND (NOT (Data[26] OR Data[47])))) AND (((NOT ((Data[16] XOR Data[7]) XOR Data[43])) OR (NOT ((FALSE XOR Data[28]) XOR Data[46]))) AND (((NOT ((Data[21] XOR Data[34]) XOR Data[39])) XOR (NOT (Data[26] OR Data[34]))) XOR ((Data[1] AND Data[44]) AND ((Data[43] XOR Data[1]) XOR Data[47]))))) XOR (((NOT (NOT Data[32])) OR (NOT (Data[5] AND Data[31]))) AND (NOT (((((Data[30] XOR Data[30]) XOR Data[37]) AND (Data[13] AND Data[50])) XOR Data[42]) XOR (((Data[20] XOR Data[44]) XOR Data[30]) OR (Data[13] OR Data[32])))))) XOR Data[26]) XOR ((Data[16] OR ((Data[18] AND ((Data[38] AND Data[9]) AND ((Data[34] XOR Data[26]) XOR Data[40]))) AND ((NOT Data[18]) AND (((Data[45] XOR TRUE) XOR Data[2]) OR (NOT Data[16]))))) OR Data[35])) XOR Data[30]) XOR (((NOT (NOT (((((Data[13] AND Data[10]) XOR ((FALSE XOR Data[33]) XOR Data[21])) XOR (NOT Data[8])) XOR (((NOT Data[35]) XOR Data[35]) XOR (Data[33] OR Data[9]))) XOR (NOT (NOT Data[34]))))) OR Data[29]) OR (NOT (Data[21] OR (((((Data[25] XOR Data[33]) XOR Data[4]) AND (NOT Data[26])) AND (NOT Data[11])) AND (((Data[43] XOR (NOT Data[3])) XOR FALSE) OR (NOT (Data[22] OR Data[8])))))))) XOR (NOT Data[41]))) XOR (((NOT (((NOT (((Data[15] AND TRUE) XOR Data[6]) XOR (Data[48] AND Data[46]))) OR (NOT (Data[44] AND (Data[19] AND Data[30])))) AND ((NOT (((Data[45] AND Data[3]) XOR Data[28]) XOR (Data[47] AND Data[44]))) AND Data[20]))) OR Data[46]) OR (((Data[27] XOR (((NOT ((Data[10] OR Data[27]) OR (Data[24] OR (Data[38] OR Data[33])))) XOR (Data[37] AND (Data[7] OR (((NOT Data[46]) XOR ((Data[20] XOR Data[42]) XOR Data[46])) XOR Data[10])))) XOR (Data[15] AND (((((FALSE XOR Data[15]) XOR Data[41]) OR (Data[19] AND Data[28])) XOR (Data[25] OR (Data[48] OR Data[14]))) XOR (NOT (NOT Data[38])))))) XOR Data[9]) AND ((((NOT ((((Data[2] OR Data[41]) XOR (Data[15] AND Data[50])) XOR (Data[39] OR Data[34])) OR (((Data[50] XOR Data[15]) XOR Data[2]) OR (NOT Data[36])))) AND Data[11]) XOR (NOT ((NOT (Data[26] AND (Data[10] AND Data[45]))) AND (NOT Data[19])))) XOR ((Data[13] AND (Data[45] OR (((Data[42] OR Data[30]) XOR (Data[44] AND TRUE)) XOR (NOT Data[46])))) OR (Data[19] AND ((NOT ((Data[26] XOR Data[9]) XOR Data[43])) AND ((NOT Data[29]) OR ((Data[11] XOR Data[23]) XOR FALSE))))))))));
    OutReady := 1;
    CollectInput(RESET:=TRUE);
  END_IF;
END_PROGRAM

CONFIGURATION Config0
  RESOURCE Res0 ON PLC
    TASK task0(INTERVAL := T#20ms,PRIORITY := 0);
    PROGRAM instance0 WITH task0 : Boiler;
  END_RESOURCE
END_CONFIGURATION
